// TIA Portal V15.1 program export: 1 tag tables, 0 data types, 3 data blocks, 7 code blocks (in call order from the OBs), 3 instance data blocks

VAR_GLOBAL   // PLC tag table "IO"
   PSH_101 AT %I0.0 : Bool;   // Scrubber high pressure
   LSH_102 AT %I0.1 : Bool;   // Scrubber high level
   LSHH_103 AT %I0.2 : Bool;   // Scrubber high-high level
   BR01_Run AT %I0.3 : Bool;   // BR01 run feedback
   S1_BR01_Start AT %I0.4 : Bool;   // BR01 START push button
   BR01_Fault AT %I0.5 : Bool;   // BR01 fault (lockout)
   S3_BR01_Stop AT %I0.6 : Bool;   // BR01 STOP push button
   S0_EStopStatus AT %I1.0 : Bool;   // E-STOP status (NC1)
   S2_FaultReset AT %I1.1 : Bool;   // FAULT RESET push button
   LSL_TK01 AT %I1.2 : Bool;   // TK01 low level
   LSL_TK02 AT %I1.3 : Bool;   // TK02 low level
   BR02_Run AT %I1.4 : Bool;   // BR02 run feedback
   BR02_Fault AT %I1.5 : Bool;   // BR02 fault (lockout)
   Rfuel2_BR02_DieselMode AT %I12.0 : Bool;   // BR02 diesel mode
   S4_BR01_Auto AT %I12.1 : Bool;   // BR01 AUTO/MAN selector (closed = AUTO)
   S5_BR02_Auto AT %I12.2 : Bool;   // BR02 AUTO/MAN selector (closed = AUTO)
   S6_BR02_Start AT %I12.3 : Bool;   // BR02 START push button
   S7_BR02_Stop AT %I12.4 : Bool;   // BR02 STOP push button
   BR01_TL_Cmd AT %Q0.0 : Bool;   // BR01 heat request (TL) + H1 1st stage lamp
   BR01_TR_Cmd AT %Q0.1 : Bool;   // BR01 2nd stage (TR) + H2 2nd stage lamp
   XV_401_Cmd AT %Q0.2 : Bool;   // XV-401 Flare SV (NO)
   XV_402_Cmd AT %Q0.3 : Bool;   // XV-402 Drain SV (NC)
   XV_403_Cmd AT %Q0.4 : Bool;   // XV-403 Suction SV (NC)
   BR02_L_Cmd AT %Q0.5 : Bool;   // BR02 start (L)
   BR02_T2_Cmd AT %Q0.6 : Bool;   // BR02 high fire (T2)
   BR02_Stage1Lamp_Cmd AT %Q0.7 : Bool;   // BR02 1st stage lamp H5
   BR02_Stage2Lamp_Cmd AT %Q1.0 : Bool;   // BR02 2nd stage lamp H6
   TE_501_Raw AT %IW96 : Int;   // TK01 inlet oil temperature
   TE_502_Raw AT %IW98 : Int;   // TK01 outlet oil temperature
   TE_503_Raw AT %IW100 : Int;   // TK02 inlet oil temperature
   TE_504_Raw AT %IW102 : Int;   // TK02 outlet oil temperature
END_VAR

DATA_BLOCK "HmiAlm"   // DB6
{ S7_Optimized_Access := 'TRUE' }
VERSION : 0.1
// stored: AutoNumber false, MemoryReserve 100
   VAR
      Common : Word;   // 0007 / H-05: x0 E-STOP active or not reset [C01]; x1 Scrubber trip: high pressure PSH-101 [C03 / C06a (PH proposal: cause memory)]; x2 Scrubber trip: high-high level LSHH-103 [C05 / C06a (PH proposal: cause memory)]; x3 Scrubber held after power-up: RESET required [S-01 / C06a (PH proposal)]; x4 Scrubber high level LSH-102 [C04 (Client)]; x5 Setting rejected: out of range [R-11]; x6 Scrubber drain open too long: drain closed [C04a]; x7 LSH-102 fault: LSHH-103 without LSH-102 [C04b]
      BR01 : Word;   // 0007 / H-05: x0 BR01 stopped by E-STOP: RESET + START [C01]; x1 BR01 thermocouple fault [C07d]; x2 BR01 burner lockout [C07e]; x3 BR01 failed to start [C07f]; x4 BR01 stopped by itself [C07g]; x5 BR01 RUN without request [R-09]; x6 TK01 level low: burner held [C07a (PH proposal: alarm; Client: permissive)]
      BR02 : Word;   // 0007 / H-05: x0 BR02 stopped by E-STOP: RESET + START [C01]; x1 BR02 thermocouple fault [C08d]; x2 BR02 burner lockout [C08e]; x3 BR02 failed to start [C08f]; x4 BR02 stopped by itself [C08g]; x5 BR02 RUN without request [R-09]; x6 TK02 level low: burner held [C08a (PH proposal: alarm; Client: permissive)]
   END_VAR
BEGIN
END_DATA_BLOCK

DATA_BLOCK "Par"   // DB1
{ S7_Optimized_Access := 'TRUE' }
VERSION : 0.1
// stored: AutoNumber false, MemoryReserve 100
   VAR RETAIN
      SP : Int := 700;   // HMI entry: Setpoint, 0.1 degC (C07b)
      HYST : Int := 50;   // HMI entry: Restart hysteresis, 0.1 degC (C07b)
      STG : Int := 100;   // HMI entry: 2nd stage below SP - STG, 0.1 degC (C07c)
      TStart : Time := T#2M;   // HMI entry: Max. time heat request -> RUN (C07f)
      TDrnOn : Time := T#3S;   // HMI entry: Scrubber high level before drain opens (C04)
      TDrnOff : Time := T#5S;   // HMI entry: Scrubber level gone before drain closes (C04)
      TDrnMax : Time := T#10M;   // HMI entry: Scrubber drain max. continuous open time (C04a)
      SP_V : Int := 700;   // Validated value used by the program (R-11)
      HYST_V : Int := 50;   // Validated value used by the program (R-11)
      STG_V : Int := 100;   // Validated value used by the program (R-11)
      TStart_V : Time := T#2M;   // Validated value used by the program (R-11)
      TDrnOn_V : Time := T#3S;   // Validated value used by the program (R-11)
      TDrnOff_V : Time := T#5S;   // Validated value used by the program (R-11)
      TDrnMax_V : Time := T#10M;   // Validated value used by the program (R-11)
   END_VAR
BEGIN
END_DATA_BLOCK

DATA_BLOCK "Sys"   // DB2
{ S7_Optimized_Access := 'TRUE' }
VERSION : 0.1
// stored: AutoNumber false, MemoryReserve 100
   VAR
      FirstScan : Bool;   // Set by OB100, cleared at the end of Main (C02)
      EStopOK : Bool;   // E-STOP latch: 1 = released and RESET given (C01)
      ResetPulse : Bool;   // RESET S2 rising edge, one scan (R-06)
      ResetMem : Bool;   // RESET edge memory (R-06)
      Alm_EStop : Bool;   // HMI alarm: E-STOP (C01)
      Alm_ParRejected : Bool;   // HMI alarm: a parameter entry was out of range (R-11)
   END_VAR
BEGIN
END_DATA_BLOCK

ORGANIZATION_BLOCK "Main"   // OB1, LAD, ProgramCycle
TITLE = Main
{ S7_Optimized_Access := 'TRUE' }
VERSION : 0.1
// Calls the blocks in a fixed order; no logic here (decisions/0006)
// stored: AutoNumber false, IsIECCheckEnabled false, SetENOAutomatically False
   VAR_INPUT
      Initial_Call : Bool;
      Remanence : Bool;
   END_VAR
BEGIN

REGION Network 1: decisions/0006 — Common: E-STOP latch, RESET edge, parameters
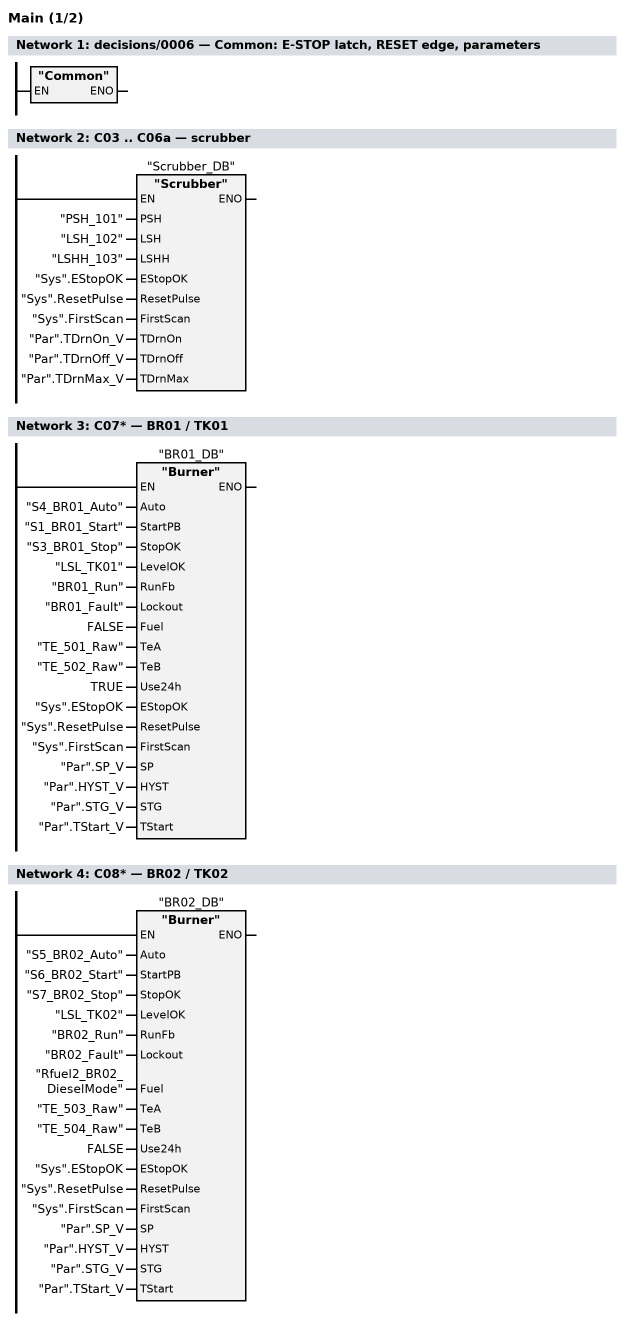
   RUNG wire#powerrail
      "Common"()
   END_RUNG
   // the same network as SCL:
   "Common"();
END_REGION

REGION Network 2: C03 .. C06a — scrubber
   RUNG wire#powerrail
      "Scrubber_DB"(PSH := "PSH_101", LSH := "LSH_102", LSHH := "LSHH_103", EStopOK := "Sys".EStopOK, ResetPulse := "Sys".ResetPulse, FirstScan := "Sys".FirstScan, TDrnOn := "Par".TDrnOn_V, TDrnOff := "Par".TDrnOff_V, TDrnMax := "Par".TDrnMax_V)
   END_RUNG
   // the same network as SCL:
   "Scrubber_DB"(PSH := "PSH_101",   // "Scrubber"
                 LSH := "LSH_102",
                 LSHH := "LSHH_103",
                 EStopOK := "Sys".EStopOK,
                 ResetPulse := "Sys".ResetPulse,
                 FirstScan := "Sys".FirstScan,
                 TDrnOn := "Par".TDrnOn_V,
                 TDrnOff := "Par".TDrnOff_V,
                 TDrnMax := "Par".TDrnMax_V);
END_REGION

REGION Network 3: C07* — BR01 / TK01
   RUNG wire#powerrail
      "BR01_DB"(Auto := "S4_BR01_Auto", StartPB := "S1_BR01_Start", StopOK := "S3_BR01_Stop", LevelOK := "LSL_TK01", RunFb := "BR01_Run", Lockout := "BR01_Fault", Fuel := FALSE, TeA := "TE_501_Raw", TeB := "TE_502_Raw", Use24h := TRUE, EStopOK := "Sys".EStopOK, ResetPulse := "Sys".ResetPulse, FirstScan := "Sys".FirstScan, SP := "Par".SP_V, HYST := "Par".HYST_V, STG := "Par".STG_V, TStart := "Par".TStart_V)
   END_RUNG
   // the same network as SCL:
   "BR01_DB"(Auto := "S4_BR01_Auto",   // "Burner"
             StartPB := "S1_BR01_Start",
             StopOK := "S3_BR01_Stop",
             LevelOK := "LSL_TK01",
             RunFb := "BR01_Run",
             Lockout := "BR01_Fault",
             Fuel := FALSE,
             TeA := "TE_501_Raw",
             TeB := "TE_502_Raw",
             Use24h := TRUE,
             EStopOK := "Sys".EStopOK,
             ResetPulse := "Sys".ResetPulse,
             FirstScan := "Sys".FirstScan,
             SP := "Par".SP_V,
             HYST := "Par".HYST_V,
             STG := "Par".STG_V,
             TStart := "Par".TStart_V);
END_REGION

REGION Network 4: C08* — BR02 / TK02
   RUNG wire#powerrail
      "BR02_DB"(Auto := "S5_BR02_Auto", StartPB := "S6_BR02_Start", StopOK := "S7_BR02_Stop", LevelOK := "LSL_TK02", RunFb := "BR02_Run", Lockout := "BR02_Fault", Fuel := "Rfuel2_BR02_DieselMode", TeA := "TE_503_Raw", TeB := "TE_504_Raw", Use24h := FALSE, EStopOK := "Sys".EStopOK, ResetPulse := "Sys".ResetPulse, FirstScan := "Sys".FirstScan, SP := "Par".SP_V, HYST := "Par".HYST_V, STG := "Par".STG_V, TStart := "Par".TStart_V)
   END_RUNG
   // the same network as SCL:
   "BR02_DB"(Auto := "S5_BR02_Auto",   // "Burner"
             StartPB := "S6_BR02_Start",
             StopOK := "S7_BR02_Stop",
             LevelOK := "LSL_TK02",
             RunFb := "BR02_Run",
             Lockout := "BR02_Fault",
             Fuel := "Rfuel2_BR02_DieselMode",
             TeA := "TE_503_Raw",
             TeB := "TE_504_Raw",
             Use24h := FALSE,
             EStopOK := "Sys".EStopOK,
             ResetPulse := "Sys".ResetPulse,
             FirstScan := "Sys".FirstScan,
             SP := "Par".SP_V,
             HYST := "Par".HYST_V,
             STG := "Par".STG_V,
             TStart := "Par".TStart_V);
END_REGION

REGION Network 5: E1 .. E7 — outputs
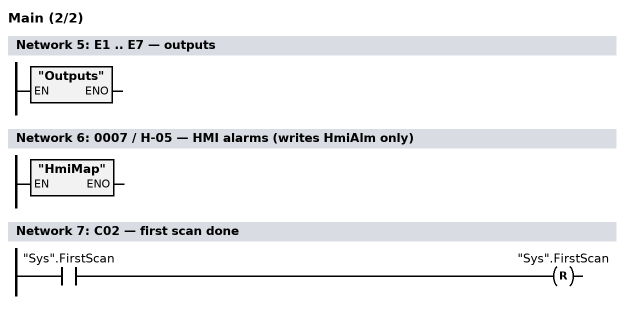
   RUNG wire#powerrail
      "Outputs"()
   END_RUNG
   // the same network as SCL:
   "Outputs"();
END_REGION

REGION Network 6: 0007 / H-05 — HMI alarms (writes HmiAlm only)
   RUNG wire#powerrail
      "HmiMap"()
   END_RUNG
   // the same network as SCL:
   "HmiMap"();
END_REGION

REGION Network 7: C02 — first scan done
   RUNG wire#powerrail
      Contact( "Sys".FirstScan )
      R_Coil( "Sys".FirstScan )
   END_RUNG
   // the same network as SCL:
   IF "Sys".FirstScan THEN "Sys".FirstScan := FALSE; END_IF;
END_REGION
END_ORGANIZATION_BLOCK

FUNCTION "Common" : Void   // FC1, LAD
TITLE = Common
{ S7_Optimized_Access := 'TRUE' }
VERSION : 0.1
// E-STOP latch, RESET edge, parameter check (decisions/0006)
// stored: AutoNumber false, IsIECCheckEnabled false, SetENOAutomatically False
   VAR_TEMP   // added for the SCL form of the ladder/FBD networks
      _w1 : Bool;
   END_VAR
BEGIN

REGION Network 1: R-06 — RESET edge (not on first scan)
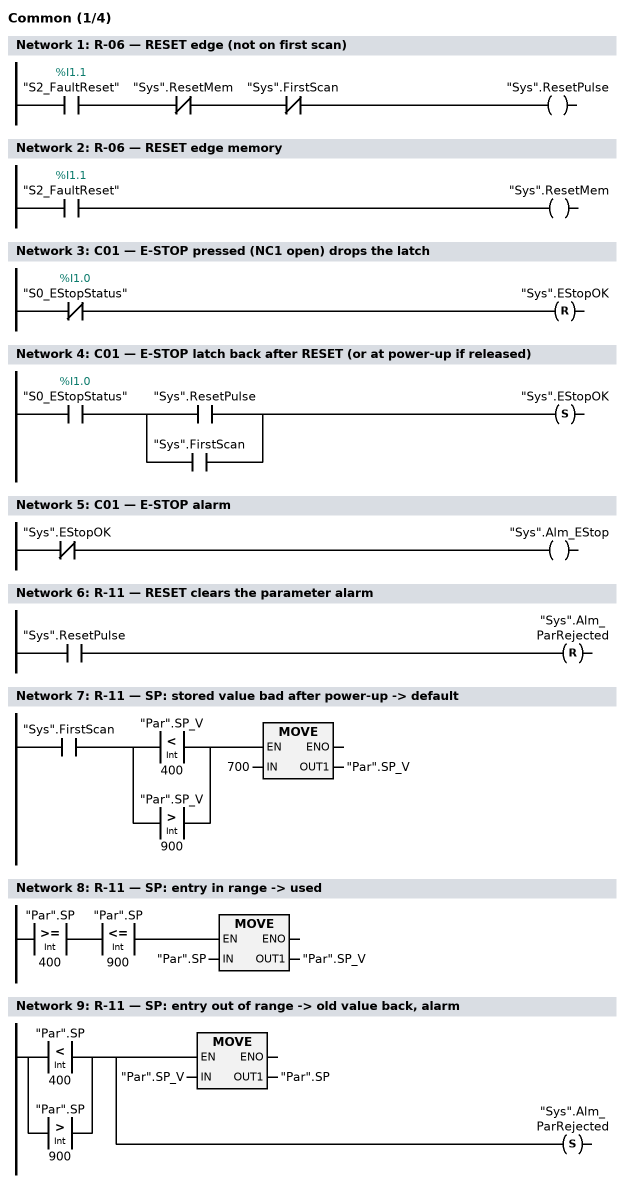
   RUNG wire#powerrail
      Contact( "S2_FaultReset" )
      I_Contact( "Sys".ResetMem )
      I_Contact( "Sys".FirstScan )
      Coil( "Sys".ResetPulse )
   END_RUNG
   // the same network as SCL:
   "Sys".ResetPulse := "S2_FaultReset" AND NOT "Sys".ResetMem AND NOT "Sys".FirstScan;
END_REGION

REGION Network 2: R-06 — RESET edge memory
   RUNG wire#powerrail
      Contact( "S2_FaultReset" )
      Coil( "Sys".ResetMem )
   END_RUNG
   // the same network as SCL:
   "Sys".ResetMem := "S2_FaultReset";
END_REGION

REGION Network 3: C01 — E-STOP pressed (NC1 open) drops the latch
   RUNG wire#powerrail
      I_Contact( "S0_EStopStatus" )
      R_Coil( "Sys".EStopOK )
   END_RUNG
   // the same network as SCL:
   IF NOT "S0_EStopStatus" THEN "Sys".EStopOK := FALSE; END_IF;
END_REGION

REGION Network 4: C01 — E-STOP latch back after RESET (or at power-up if released)
   RUNG wire#powerrail
      Contact( "S0_EStopStatus" )
      wire#w1
      Contact( "Sys".ResetPulse )
      wire#w2
      S_Coil( "Sys".EStopOK )
   END_RUNG
   RUNG wire#w1
      Contact( "Sys".FirstScan )
   END_RUNG wire#w2
   // the same network as SCL:
   IF "S0_EStopStatus" AND ("Sys".ResetPulse OR "Sys".FirstScan) THEN "Sys".EStopOK := TRUE; END_IF;
END_REGION

REGION Network 5: C01 — E-STOP alarm
   RUNG wire#powerrail
      I_Contact( "Sys".EStopOK )
      Coil( "Sys".Alm_EStop )
   END_RUNG
   // the same network as SCL:
   "Sys".Alm_EStop := NOT "Sys".EStopOK;
END_REGION

REGION Network 6: R-11 — RESET clears the parameter alarm
   RUNG wire#powerrail
      Contact( "Sys".ResetPulse )
      R_Coil( "Sys".Alm_ParRejected )
   END_RUNG
   // the same network as SCL:
   IF "Sys".ResetPulse THEN "Sys".Alm_ParRejected := FALSE; END_IF;
END_REGION

REGION Network 7: R-11 — SP: stored value bad after power-up -> default
   RUNG wire#powerrail
      Contact( "Sys".FirstScan )
      wire#w1
      { S7_Templates := "SrcType := Int" } LT_Contact(in1 := "Par".SP_V, in2 := 400)
      wire#w2
      { S7_GenerateENO := "TRUE" } Move(in := 700, out1 => "Par".SP_V)
   END_RUNG
   RUNG wire#w1
      { S7_Templates := "SrcType := Int" } GT_Contact(in1 := "Par".SP_V, in2 := 900)
   END_RUNG wire#w2
   // the same network as SCL:
   IF "Sys".FirstScan AND (("Par".SP_V < 400) OR ("Par".SP_V > 900)) THEN "Par".SP_V := 700; END_IF;
END_REGION

REGION Network 8: R-11 — SP: entry in range -> used
   RUNG wire#powerrail
      { S7_Templates := "SrcType := Int" } GE_Contact(in1 := "Par".SP, in2 := 400)
      { S7_Templates := "SrcType := Int" } LE_Contact(in1 := "Par".SP, in2 := 900)
      { S7_GenerateENO := "TRUE" } Move(in := "Par".SP, out1 => "Par".SP_V)
   END_RUNG
   // the same network as SCL:
   IF ("Par".SP >= 400) AND ("Par".SP <= 900) THEN "Par".SP_V := "Par".SP; END_IF;
END_REGION

REGION Network 9: R-11 — SP: entry out of range -> old value back, alarm
   RUNG wire#powerrail
      { S7_Templates := "SrcType := Int" } LT_Contact(in1 := "Par".SP, in2 := 400)
      wire#w1
      { S7_GenerateENO := "TRUE" } Move(in := "Par".SP_V, out1 => "Par".SP)
   END_RUNG
   RUNG wire#powerrail
      { S7_Templates := "SrcType := Int" } GT_Contact(in1 := "Par".SP, in2 := 900)
   END_RUNG wire#w1
   RUNG wire#w1
      S_Coil( "Sys".Alm_ParRejected )
   END_RUNG
   // the same network as SCL:
   #_w1 := ("Par".SP < 400) OR ("Par".SP > 900);
   IF #_w1 THEN
       "Par".SP := "Par".SP_V;
       "Sys".Alm_ParRejected := TRUE;
   END_IF;
END_REGION

REGION Network 10: R-11 — HYST: stored value bad after power-up -> default
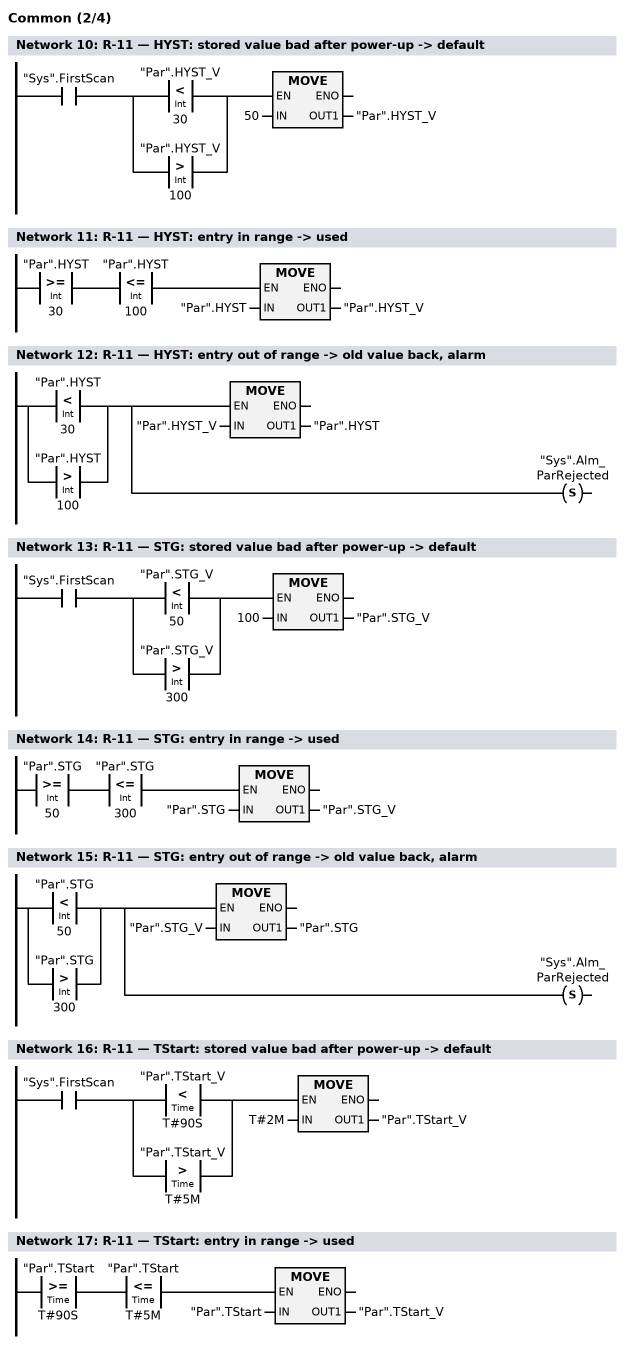
   RUNG wire#powerrail
      Contact( "Sys".FirstScan )
      wire#w1
      { S7_Templates := "SrcType := Int" } LT_Contact(in1 := "Par".HYST_V, in2 := 30)
      wire#w2
      { S7_GenerateENO := "TRUE" } Move(in := 50, out1 => "Par".HYST_V)
   END_RUNG
   RUNG wire#w1
      { S7_Templates := "SrcType := Int" } GT_Contact(in1 := "Par".HYST_V, in2 := 100)
   END_RUNG wire#w2
   // the same network as SCL:
   IF "Sys".FirstScan AND (("Par".HYST_V < 30) OR ("Par".HYST_V > 100)) THEN "Par".HYST_V := 50; END_IF;
END_REGION

REGION Network 11: R-11 — HYST: entry in range -> used
   RUNG wire#powerrail
      { S7_Templates := "SrcType := Int" } GE_Contact(in1 := "Par".HYST, in2 := 30)
      { S7_Templates := "SrcType := Int" } LE_Contact(in1 := "Par".HYST, in2 := 100)
      { S7_GenerateENO := "TRUE" } Move(in := "Par".HYST, out1 => "Par".HYST_V)
   END_RUNG
   // the same network as SCL:
   IF ("Par".HYST >= 30) AND ("Par".HYST <= 100) THEN "Par".HYST_V := "Par".HYST; END_IF;
END_REGION

REGION Network 12: R-11 — HYST: entry out of range -> old value back, alarm
   RUNG wire#powerrail
      { S7_Templates := "SrcType := Int" } LT_Contact(in1 := "Par".HYST, in2 := 30)
      wire#w1
      { S7_GenerateENO := "TRUE" } Move(in := "Par".HYST_V, out1 => "Par".HYST)
   END_RUNG
   RUNG wire#powerrail
      { S7_Templates := "SrcType := Int" } GT_Contact(in1 := "Par".HYST, in2 := 100)
   END_RUNG wire#w1
   RUNG wire#w1
      S_Coil( "Sys".Alm_ParRejected )
   END_RUNG
   // the same network as SCL:
   #_w1 := ("Par".HYST < 30) OR ("Par".HYST > 100);
   IF #_w1 THEN
       "Par".HYST := "Par".HYST_V;
       "Sys".Alm_ParRejected := TRUE;
   END_IF;
END_REGION

REGION Network 13: R-11 — STG: stored value bad after power-up -> default
   RUNG wire#powerrail
      Contact( "Sys".FirstScan )
      wire#w1
      { S7_Templates := "SrcType := Int" } LT_Contact(in1 := "Par".STG_V, in2 := 50)
      wire#w2
      { S7_GenerateENO := "TRUE" } Move(in := 100, out1 => "Par".STG_V)
   END_RUNG
   RUNG wire#w1
      { S7_Templates := "SrcType := Int" } GT_Contact(in1 := "Par".STG_V, in2 := 300)
   END_RUNG wire#w2
   // the same network as SCL:
   IF "Sys".FirstScan AND (("Par".STG_V < 50) OR ("Par".STG_V > 300)) THEN "Par".STG_V := 100; END_IF;
END_REGION

REGION Network 14: R-11 — STG: entry in range -> used
   RUNG wire#powerrail
      { S7_Templates := "SrcType := Int" } GE_Contact(in1 := "Par".STG, in2 := 50)
      { S7_Templates := "SrcType := Int" } LE_Contact(in1 := "Par".STG, in2 := 300)
      { S7_GenerateENO := "TRUE" } Move(in := "Par".STG, out1 => "Par".STG_V)
   END_RUNG
   // the same network as SCL:
   IF ("Par".STG >= 50) AND ("Par".STG <= 300) THEN "Par".STG_V := "Par".STG; END_IF;
END_REGION

REGION Network 15: R-11 — STG: entry out of range -> old value back, alarm
   RUNG wire#powerrail
      { S7_Templates := "SrcType := Int" } LT_Contact(in1 := "Par".STG, in2 := 50)
      wire#w1
      { S7_GenerateENO := "TRUE" } Move(in := "Par".STG_V, out1 => "Par".STG)
   END_RUNG
   RUNG wire#powerrail
      { S7_Templates := "SrcType := Int" } GT_Contact(in1 := "Par".STG, in2 := 300)
   END_RUNG wire#w1
   RUNG wire#w1
      S_Coil( "Sys".Alm_ParRejected )
   END_RUNG
   // the same network as SCL:
   #_w1 := ("Par".STG < 50) OR ("Par".STG > 300);
   IF #_w1 THEN
       "Par".STG := "Par".STG_V;
       "Sys".Alm_ParRejected := TRUE;
   END_IF;
END_REGION

REGION Network 16: R-11 — TStart: stored value bad after power-up -> default
   RUNG wire#powerrail
      Contact( "Sys".FirstScan )
      wire#w1
      { S7_Templates := "SrcType := Time" } LT_Contact(in1 := "Par".TStart_V, in2 := T#90S)
      wire#w2
      { S7_GenerateENO := "TRUE" } Move(in := T#2M, out1 => "Par".TStart_V)
   END_RUNG
   RUNG wire#w1
      { S7_Templates := "SrcType := Time" } GT_Contact(in1 := "Par".TStart_V, in2 := T#5M)
   END_RUNG wire#w2
   // the same network as SCL:
   IF "Sys".FirstScan AND (("Par".TStart_V < T#90S) OR ("Par".TStart_V > T#5M)) THEN
       "Par".TStart_V := T#2M;
   END_IF;
END_REGION

REGION Network 17: R-11 — TStart: entry in range -> used
   RUNG wire#powerrail
      { S7_Templates := "SrcType := Time" } GE_Contact(in1 := "Par".TStart, in2 := T#90S)
      { S7_Templates := "SrcType := Time" } LE_Contact(in1 := "Par".TStart, in2 := T#5M)
      { S7_GenerateENO := "TRUE" } Move(in := "Par".TStart, out1 => "Par".TStart_V)
   END_RUNG
   // the same network as SCL:
   IF ("Par".TStart >= T#90S) AND ("Par".TStart <= T#5M) THEN "Par".TStart_V := "Par".TStart; END_IF;
END_REGION

REGION Network 18: R-11 — TStart: entry out of range -> old value back, alarm
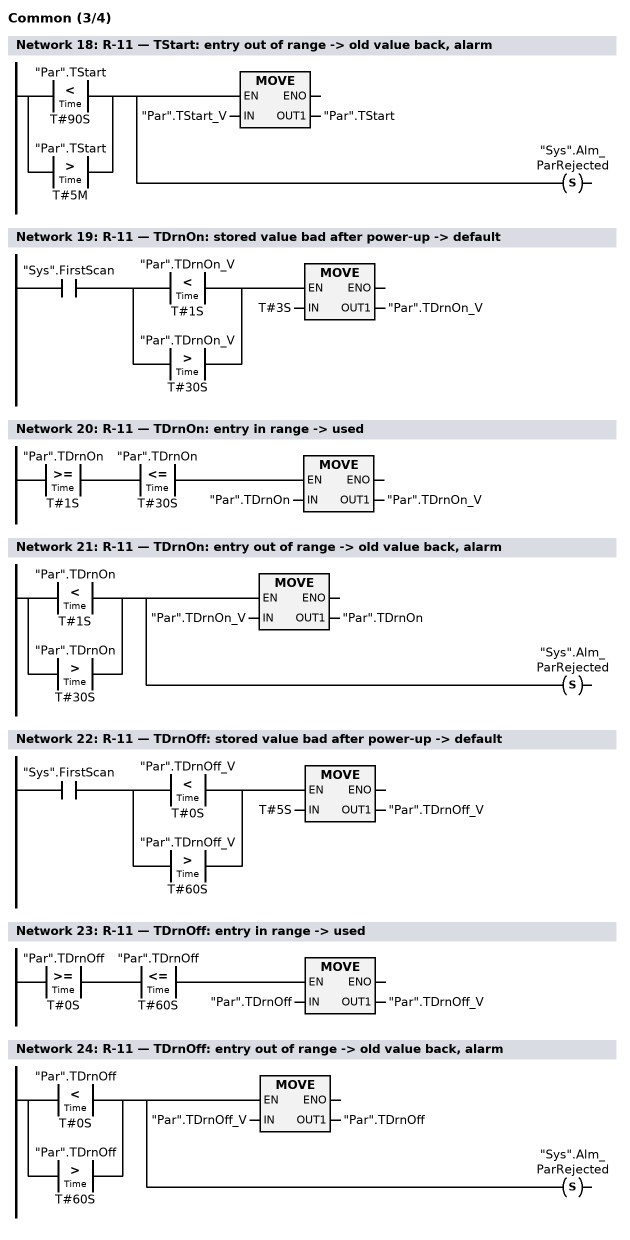
   RUNG wire#powerrail
      { S7_Templates := "SrcType := Time" } LT_Contact(in1 := "Par".TStart, in2 := T#90S)
      wire#w1
      { S7_GenerateENO := "TRUE" } Move(in := "Par".TStart_V, out1 => "Par".TStart)
   END_RUNG
   RUNG wire#powerrail
      { S7_Templates := "SrcType := Time" } GT_Contact(in1 := "Par".TStart, in2 := T#5M)
   END_RUNG wire#w1
   RUNG wire#w1
      S_Coil( "Sys".Alm_ParRejected )
   END_RUNG
   // the same network as SCL:
   #_w1 := ("Par".TStart < T#90S) OR ("Par".TStart > T#5M);
   IF #_w1 THEN
       "Par".TStart := "Par".TStart_V;
       "Sys".Alm_ParRejected := TRUE;
   END_IF;
END_REGION

REGION Network 19: R-11 — TDrnOn: stored value bad after power-up -> default
   RUNG wire#powerrail
      Contact( "Sys".FirstScan )
      wire#w1
      { S7_Templates := "SrcType := Time" } LT_Contact(in1 := "Par".TDrnOn_V, in2 := T#1S)
      wire#w2
      { S7_GenerateENO := "TRUE" } Move(in := T#3S, out1 => "Par".TDrnOn_V)
   END_RUNG
   RUNG wire#w1
      { S7_Templates := "SrcType := Time" } GT_Contact(in1 := "Par".TDrnOn_V, in2 := T#30S)
   END_RUNG wire#w2
   // the same network as SCL:
   IF "Sys".FirstScan AND (("Par".TDrnOn_V < T#1S) OR ("Par".TDrnOn_V > T#30S)) THEN
       "Par".TDrnOn_V := T#3S;
   END_IF;
END_REGION

REGION Network 20: R-11 — TDrnOn: entry in range -> used
   RUNG wire#powerrail
      { S7_Templates := "SrcType := Time" } GE_Contact(in1 := "Par".TDrnOn, in2 := T#1S)
      { S7_Templates := "SrcType := Time" } LE_Contact(in1 := "Par".TDrnOn, in2 := T#30S)
      { S7_GenerateENO := "TRUE" } Move(in := "Par".TDrnOn, out1 => "Par".TDrnOn_V)
   END_RUNG
   // the same network as SCL:
   IF ("Par".TDrnOn >= T#1S) AND ("Par".TDrnOn <= T#30S) THEN "Par".TDrnOn_V := "Par".TDrnOn; END_IF;
END_REGION

REGION Network 21: R-11 — TDrnOn: entry out of range -> old value back, alarm
   RUNG wire#powerrail
      { S7_Templates := "SrcType := Time" } LT_Contact(in1 := "Par".TDrnOn, in2 := T#1S)
      wire#w1
      { S7_GenerateENO := "TRUE" } Move(in := "Par".TDrnOn_V, out1 => "Par".TDrnOn)
   END_RUNG
   RUNG wire#powerrail
      { S7_Templates := "SrcType := Time" } GT_Contact(in1 := "Par".TDrnOn, in2 := T#30S)
   END_RUNG wire#w1
   RUNG wire#w1
      S_Coil( "Sys".Alm_ParRejected )
   END_RUNG
   // the same network as SCL:
   #_w1 := ("Par".TDrnOn < T#1S) OR ("Par".TDrnOn > T#30S);
   IF #_w1 THEN
       "Par".TDrnOn := "Par".TDrnOn_V;
       "Sys".Alm_ParRejected := TRUE;
   END_IF;
END_REGION

REGION Network 22: R-11 — TDrnOff: stored value bad after power-up -> default
   RUNG wire#powerrail
      Contact( "Sys".FirstScan )
      wire#w1
      { S7_Templates := "SrcType := Time" } LT_Contact(in1 := "Par".TDrnOff_V, in2 := T#0S)
      wire#w2
      { S7_GenerateENO := "TRUE" } Move(in := T#5S, out1 => "Par".TDrnOff_V)
   END_RUNG
   RUNG wire#w1
      { S7_Templates := "SrcType := Time" } GT_Contact(in1 := "Par".TDrnOff_V, in2 := T#60S)
   END_RUNG wire#w2
   // the same network as SCL:
   IF "Sys".FirstScan AND (("Par".TDrnOff_V < T#0S) OR ("Par".TDrnOff_V > T#60S)) THEN
       "Par".TDrnOff_V := T#5S;
   END_IF;
END_REGION

REGION Network 23: R-11 — TDrnOff: entry in range -> used
   RUNG wire#powerrail
      { S7_Templates := "SrcType := Time" } GE_Contact(in1 := "Par".TDrnOff, in2 := T#0S)
      { S7_Templates := "SrcType := Time" } LE_Contact(in1 := "Par".TDrnOff, in2 := T#60S)
      { S7_GenerateENO := "TRUE" } Move(in := "Par".TDrnOff, out1 => "Par".TDrnOff_V)
   END_RUNG
   // the same network as SCL:
   IF ("Par".TDrnOff >= T#0S) AND ("Par".TDrnOff <= T#60S) THEN "Par".TDrnOff_V := "Par".TDrnOff; END_IF;
END_REGION

REGION Network 24: R-11 — TDrnOff: entry out of range -> old value back, alarm
   RUNG wire#powerrail
      { S7_Templates := "SrcType := Time" } LT_Contact(in1 := "Par".TDrnOff, in2 := T#0S)
      wire#w1
      { S7_GenerateENO := "TRUE" } Move(in := "Par".TDrnOff_V, out1 => "Par".TDrnOff)
   END_RUNG
   RUNG wire#powerrail
      { S7_Templates := "SrcType := Time" } GT_Contact(in1 := "Par".TDrnOff, in2 := T#60S)
   END_RUNG wire#w1
   RUNG wire#w1
      S_Coil( "Sys".Alm_ParRejected )
   END_RUNG
   // the same network as SCL:
   #_w1 := ("Par".TDrnOff < T#0S) OR ("Par".TDrnOff > T#60S);
   IF #_w1 THEN
       "Par".TDrnOff := "Par".TDrnOff_V;
       "Sys".Alm_ParRejected := TRUE;
   END_IF;
END_REGION

REGION Network 25: R-11 — TDrnMax: stored value bad after power-up -> default
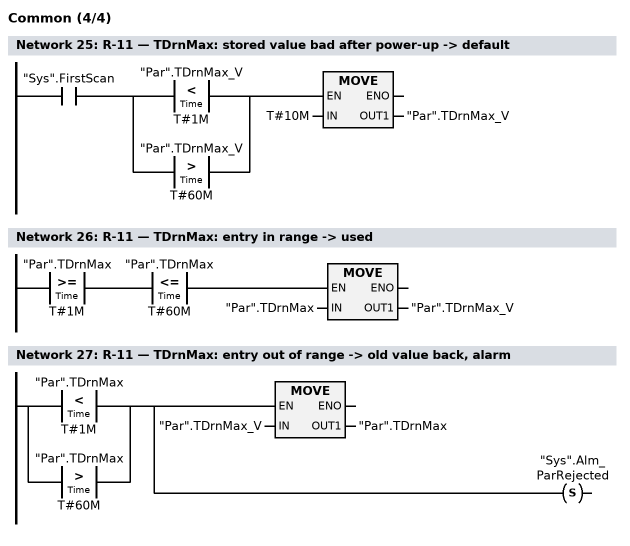
   RUNG wire#powerrail
      Contact( "Sys".FirstScan )
      wire#w1
      { S7_Templates := "SrcType := Time" } LT_Contact(in1 := "Par".TDrnMax_V, in2 := T#1M)
      wire#w2
      { S7_GenerateENO := "TRUE" } Move(in := T#10M, out1 => "Par".TDrnMax_V)
   END_RUNG
   RUNG wire#w1
      { S7_Templates := "SrcType := Time" } GT_Contact(in1 := "Par".TDrnMax_V, in2 := T#60M)
   END_RUNG wire#w2
   // the same network as SCL:
   IF "Sys".FirstScan AND (("Par".TDrnMax_V < T#1M) OR ("Par".TDrnMax_V > T#60M)) THEN
       "Par".TDrnMax_V := T#10M;
   END_IF;
END_REGION

REGION Network 26: R-11 — TDrnMax: entry in range -> used
   RUNG wire#powerrail
      { S7_Templates := "SrcType := Time" } GE_Contact(in1 := "Par".TDrnMax, in2 := T#1M)
      { S7_Templates := "SrcType := Time" } LE_Contact(in1 := "Par".TDrnMax, in2 := T#60M)
      { S7_GenerateENO := "TRUE" } Move(in := "Par".TDrnMax, out1 => "Par".TDrnMax_V)
   END_RUNG
   // the same network as SCL:
   IF ("Par".TDrnMax >= T#1M) AND ("Par".TDrnMax <= T#60M) THEN "Par".TDrnMax_V := "Par".TDrnMax; END_IF;
END_REGION

REGION Network 27: R-11 — TDrnMax: entry out of range -> old value back, alarm
   RUNG wire#powerrail
      { S7_Templates := "SrcType := Time" } LT_Contact(in1 := "Par".TDrnMax, in2 := T#1M)
      wire#w1
      { S7_GenerateENO := "TRUE" } Move(in := "Par".TDrnMax_V, out1 => "Par".TDrnMax)
   END_RUNG
   RUNG wire#powerrail
      { S7_Templates := "SrcType := Time" } GT_Contact(in1 := "Par".TDrnMax, in2 := T#60M)
   END_RUNG wire#w1
   RUNG wire#w1
      S_Coil( "Sys".Alm_ParRejected )
   END_RUNG
   // the same network as SCL:
   #_w1 := ("Par".TDrnMax < T#1M) OR ("Par".TDrnMax > T#60M);
   IF #_w1 THEN
       "Par".TDrnMax := "Par".TDrnMax_V;
       "Sys".Alm_ParRejected := TRUE;
   END_IF;
END_REGION
END_FUNCTION

FUNCTION_BLOCK "Scrubber"   // FB2, LAD
TITLE = Scrubber
{ S7_Optimized_Access := 'TRUE' }
VERSION : 0.1
// Gas scrubber, docs/التشغيل.md §1
// stored: AutoNumber false, IsIECCheckEnabled false, MemoryReserve 100, SetENOAutomatically False
   VAR_INPUT
      PSH : Bool;   // PSH-101 healthy (contact closed)
      LSH : Bool;   // LSH-102 healthy
      LSHH : Bool;   // LSHH-103 healthy
      EStopOK : Bool;   // Sys.EStopOK
      ResetPulse : Bool;   // Sys.ResetPulse
      FirstScan : Bool;   // Sys.FirstScan
      TDrnOn : Time;   // Par.TDrnOn_V (C04)
      TDrnOff : Time;   // Par.TDrnOff_V (C04)
      TDrnMax : Time;   // Par.TDrnMax_V (C04a)
   END_VAR
   VAR_OUTPUT
      Tripped : Bool;   // Suction trip latch C01/C02/C03/C05: XV-403 closed until RESET
      FlareTrip : Bool;   // Flare trip latch C01/C02/C03: XV-401 open until RESET
      ValvesNormal : Bool;   // No trip latched: flare closed and suction open (HMI)
      FlareCmd : Bool;   // Q0.2 XV-401 (NO): 1 = energised = closed
      DrainCmd : Bool;   // Q0.3 XV-402 (NC): 1 = energised = open (C04 / C05)
      SuctionCmd : Bool;   // Q0.4 XV-403 (NC): 1 = energised = open
      F_DrainTO : Bool;   // C04a: drain open too long, latched until RESET
      F_LshFault : Bool;   // C04b: LSHH-103 without LSH-102, latched until RESET
      Alm_PSH : Bool;   // HMI alarm C03
      Alm_LSH : Bool;   // HMI alarm C04
      Alm_LSHH : Bool;   // HMI alarm C05
      Cause_EStop : Bool;   // C06a / F44: E-STOP cause, latched until healthy RESET
      Cause_PSH : Bool;   // C06a / F44: PSH-101 cause, latched until healthy RESET
      Cause_LSHH : Bool;   // C06a / F44: LSHH-103 cause, latched until healthy RESET
      Cause_PwrUp : Bool;   // C06a / F44: power-up cause, latched until healthy RESET
      FirstOut : Int;   // C06a / 0007 D5: 0 none, 1 E-STOP, 2 PSH, 3 LSHH, 4 power-up
   END_VAR
   VAR
      LevelHigh : Bool;
      DrnDemand : Bool;
      T_DrnOn : TON_TIME;
      T_DrnOff : TON_TIME;
      T_DrnMax : TON_TIME;
      T_LshFlt : TON_TIME;
   END_VAR
BEGIN

REGION Network 1: C04 — LSH-102 high level alarm
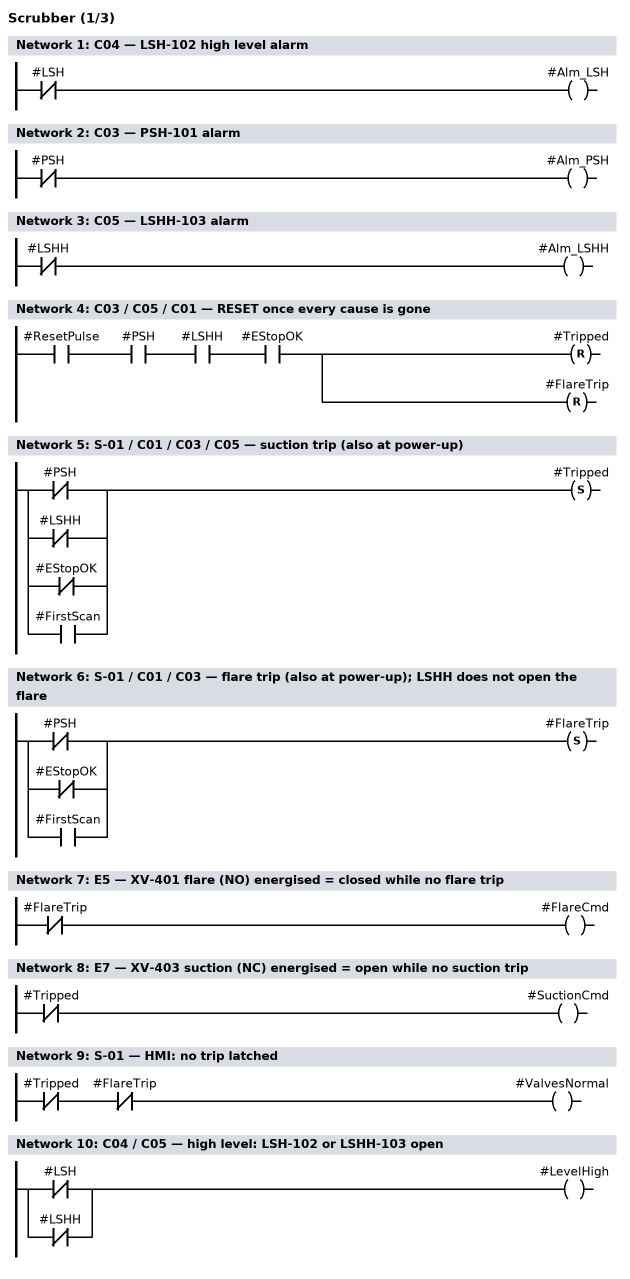
   RUNG wire#powerrail
      I_Contact( #LSH )
      Coil( #Alm_LSH )
   END_RUNG
   // the same network as SCL:
   #Alm_LSH := NOT #LSH;
END_REGION

REGION Network 2: C03 — PSH-101 alarm
   RUNG wire#powerrail
      I_Contact( #PSH )
      Coil( #Alm_PSH )
   END_RUNG
   // the same network as SCL:
   #Alm_PSH := NOT #PSH;
END_REGION

REGION Network 3: C05 — LSHH-103 alarm
   RUNG wire#powerrail
      I_Contact( #LSHH )
      Coil( #Alm_LSHH )
   END_RUNG
   // the same network as SCL:
   #Alm_LSHH := NOT #LSHH;
END_REGION

REGION Network 4: C03 / C05 / C01 — RESET once every cause is gone
   RUNG wire#powerrail
      Contact( #ResetPulse )
      Contact( #PSH )
      Contact( #LSHH )
      Contact( #EStopOK )
      wire#w1
      R_Coil( #Tripped )
   END_RUNG
   RUNG wire#w1
      R_Coil( #FlareTrip )
   END_RUNG
   // the same network as SCL:
   IF #ResetPulse AND #PSH AND #LSHH AND #EStopOK THEN
       #Tripped := FALSE;
       #FlareTrip := FALSE;
   END_IF;
END_REGION

REGION Network 5: S-01 / C01 / C03 / C05 — suction trip (also at power-up)
   RUNG wire#powerrail
      I_Contact( #PSH )
      wire#w1
      S_Coil( #Tripped )
   END_RUNG
   RUNG wire#powerrail
      I_Contact( #LSHH )
   END_RUNG wire#w1
   RUNG wire#powerrail
      I_Contact( #EStopOK )
   END_RUNG wire#w1
   RUNG wire#powerrail
      Contact( #FirstScan )
   END_RUNG wire#w1
   // the same network as SCL:
   IF NOT #PSH OR NOT #LSHH OR NOT #EStopOK OR #FirstScan THEN #Tripped := TRUE; END_IF;
END_REGION

REGION Network 6: S-01 / C01 / C03 — flare trip (also at power-up); LSHH does not open the flare
   RUNG wire#powerrail
      I_Contact( #PSH )
      wire#w1
      S_Coil( #FlareTrip )
   END_RUNG
   RUNG wire#powerrail
      I_Contact( #EStopOK )
   END_RUNG wire#w1
   RUNG wire#powerrail
      Contact( #FirstScan )
   END_RUNG wire#w1
   // the same network as SCL:
   IF NOT #PSH OR NOT #EStopOK OR #FirstScan THEN #FlareTrip := TRUE; END_IF;
END_REGION

REGION Network 7: E5 — XV-401 flare (NO) energised = closed while no flare trip
   RUNG wire#powerrail
      I_Contact( #FlareTrip )
      Coil( #FlareCmd )
   END_RUNG
   // the same network as SCL:
   #FlareCmd := NOT #FlareTrip;
END_REGION

REGION Network 8: E7 — XV-403 suction (NC) energised = open while no suction trip
   RUNG wire#powerrail
      I_Contact( #Tripped )
      Coil( #SuctionCmd )
   END_RUNG
   // the same network as SCL:
   #SuctionCmd := NOT #Tripped;
END_REGION

REGION Network 9: S-01 — HMI: no trip latched
   RUNG wire#powerrail
      I_Contact( #Tripped )
      I_Contact( #FlareTrip )
      Coil( #ValvesNormal )
   END_RUNG
   // the same network as SCL:
   #ValvesNormal := NOT #Tripped AND NOT #FlareTrip;
END_REGION

REGION Network 10: C04 / C05 — high level: LSH-102 or LSHH-103 open
   RUNG wire#powerrail
      I_Contact( #LSH )
      wire#w1
      Coil( #LevelHigh )
   END_RUNG
   RUNG wire#powerrail
      I_Contact( #LSHH )
   END_RUNG wire#w1
   // the same network as SCL:
   #LevelHigh := NOT #LSH OR NOT #LSHH;
END_REGION

REGION Network 11: C04 — drain demand after TDRN_ON of high level
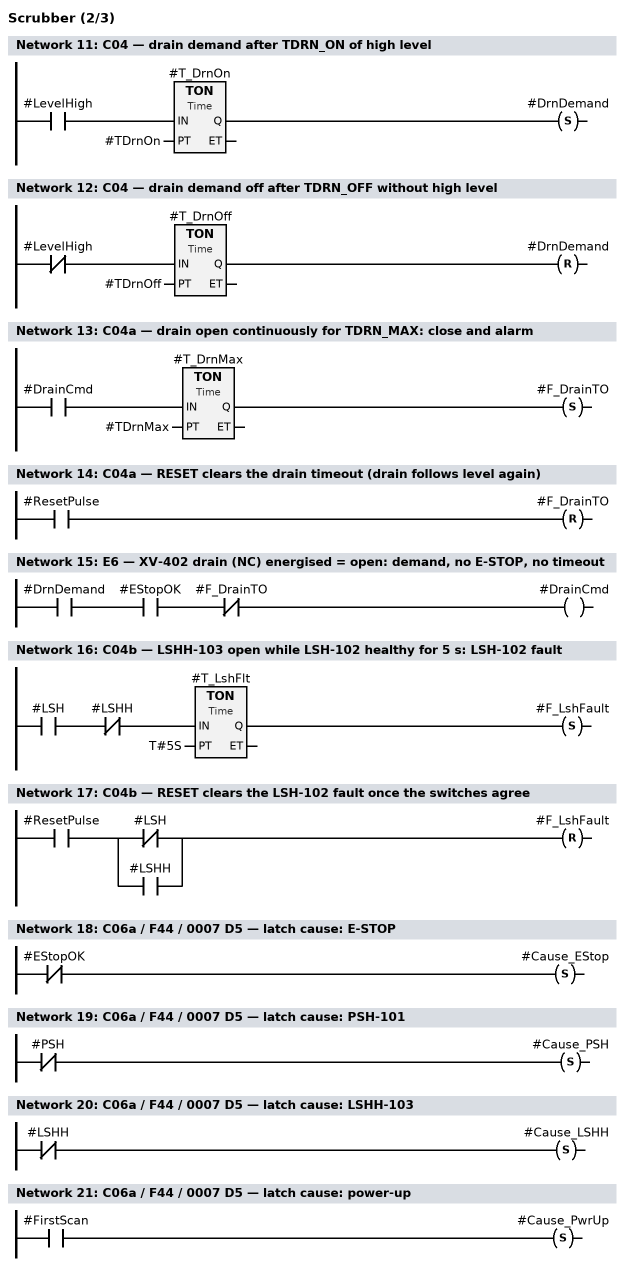
   RUNG wire#powerrail
      Contact( #LevelHigh )
      { S7_Templates := "time_type := Time" } #T_DrnOn.TON(pt := #TDrnOn, et =>)
      S_Coil( #DrnDemand )
   END_RUNG
   // the same network as SCL:
   #T_DrnOn(IN := #LevelHigh, PT := #TDrnOn);   // TON
   IF #T_DrnOn.Q THEN #DrnDemand := TRUE; END_IF;
END_REGION

REGION Network 12: C04 — drain demand off after TDRN_OFF without high level
   RUNG wire#powerrail
      I_Contact( #LevelHigh )
      { S7_Templates := "time_type := Time" } #T_DrnOff.TON(pt := #TDrnOff, et =>)
      R_Coil( #DrnDemand )
   END_RUNG
   // the same network as SCL:
   #T_DrnOff(IN := NOT #LevelHigh, PT := #TDrnOff);   // TON
   IF #T_DrnOff.Q THEN #DrnDemand := FALSE; END_IF;
END_REGION

REGION Network 13: C04a — drain open continuously for TDRN_MAX: close and alarm
   RUNG wire#powerrail
      Contact( #DrainCmd )
      { S7_Templates := "time_type := Time" } #T_DrnMax.TON(pt := #TDrnMax, et =>)
      S_Coil( #F_DrainTO )
   END_RUNG
   // the same network as SCL:
   #T_DrnMax(IN := #DrainCmd, PT := #TDrnMax);   // TON
   IF #T_DrnMax.Q THEN #F_DrainTO := TRUE; END_IF;
END_REGION

REGION Network 14: C04a — RESET clears the drain timeout (drain follows level again)
   RUNG wire#powerrail
      Contact( #ResetPulse )
      R_Coil( #F_DrainTO )
   END_RUNG
   // the same network as SCL:
   IF #ResetPulse THEN #F_DrainTO := FALSE; END_IF;
END_REGION

REGION Network 15: E6 — XV-402 drain (NC) energised = open: demand, no E-STOP, no timeout
   RUNG wire#powerrail
      Contact( #DrnDemand )
      Contact( #EStopOK )
      I_Contact( #F_DrainTO )
      Coil( #DrainCmd )
   END_RUNG
   // the same network as SCL:
   #DrainCmd := #DrnDemand AND #EStopOK AND NOT #F_DrainTO;
END_REGION

REGION Network 16: C04b — LSHH-103 open while LSH-102 healthy for 5 s: LSH-102 fault
   RUNG wire#powerrail
      Contact( #LSH )
      I_Contact( #LSHH )
      { S7_Templates := "time_type := Time" } #T_LshFlt.TON(pt := T#5S, et =>)
      S_Coil( #F_LshFault )
   END_RUNG
   // the same network as SCL:
   #T_LshFlt(IN := #LSH AND NOT #LSHH, PT := T#5S);   // TON
   IF #T_LshFlt.Q THEN #F_LshFault := TRUE; END_IF;
END_REGION

REGION Network 17: C04b — RESET clears the LSH-102 fault once the switches agree
   RUNG wire#powerrail
      Contact( #ResetPulse )
      wire#w1
      I_Contact( #LSH )
      wire#w2
      R_Coil( #F_LshFault )
   END_RUNG
   RUNG wire#w1
      Contact( #LSHH )
   END_RUNG wire#w2
   // the same network as SCL:
   IF #ResetPulse AND (NOT #LSH OR #LSHH) THEN #F_LshFault := FALSE; END_IF;
END_REGION

REGION Network 18: C06a / F44 / 0007 D5 — latch cause: E-STOP
   RUNG wire#powerrail
      I_Contact( #EStopOK )
      S_Coil( #Cause_EStop )
   END_RUNG
   // the same network as SCL:
   IF NOT #EStopOK THEN #Cause_EStop := TRUE; END_IF;
END_REGION

REGION Network 19: C06a / F44 / 0007 D5 — latch cause: PSH-101
   RUNG wire#powerrail
      I_Contact( #PSH )
      S_Coil( #Cause_PSH )
   END_RUNG
   // the same network as SCL:
   IF NOT #PSH THEN #Cause_PSH := TRUE; END_IF;
END_REGION

REGION Network 20: C06a / F44 / 0007 D5 — latch cause: LSHH-103
   RUNG wire#powerrail
      I_Contact( #LSHH )
      S_Coil( #Cause_LSHH )
   END_RUNG
   // the same network as SCL:
   IF NOT #LSHH THEN #Cause_LSHH := TRUE; END_IF;
END_REGION

REGION Network 21: C06a / F44 / 0007 D5 — latch cause: power-up
   RUNG wire#powerrail
      Contact( #FirstScan )
      S_Coil( #Cause_PwrUp )
   END_RUNG
   // the same network as SCL:
   IF #FirstScan THEN #Cause_PwrUp := TRUE; END_IF;
END_REGION

REGION Network 22: C06a / F44 / 0007 D5 — first-out 1: E-STOP (only if none)
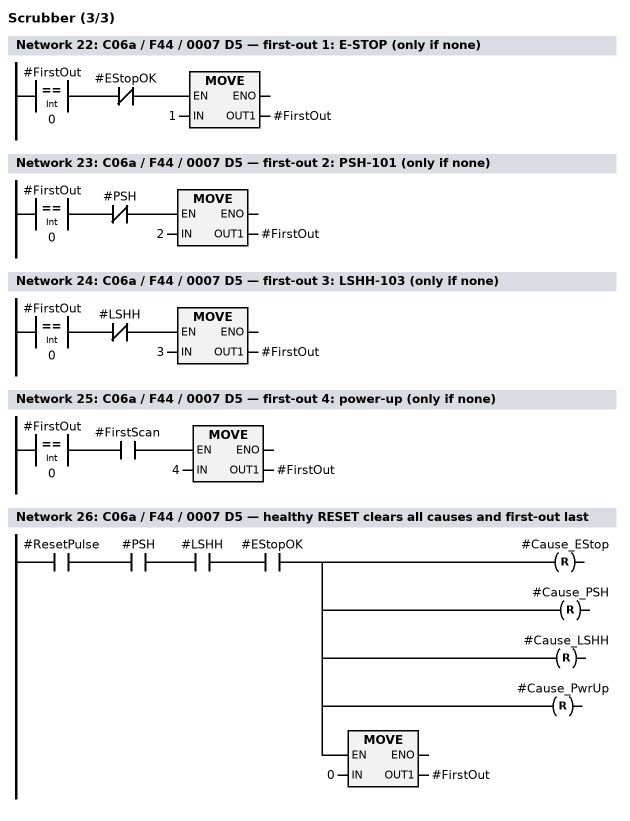
   RUNG wire#powerrail
      { S7_Templates := "SrcType := Int" } EQ_Contact(in1 := #FirstOut, in2 := 0)
      I_Contact( #EStopOK )
      { S7_GenerateENO := "TRUE" } Move(in := 1, out1 => #FirstOut)
   END_RUNG
   // the same network as SCL:
   IF (#FirstOut = 0) AND NOT #EStopOK THEN #FirstOut := 1; END_IF;
END_REGION

REGION Network 23: C06a / F44 / 0007 D5 — first-out 2: PSH-101 (only if none)
   RUNG wire#powerrail
      { S7_Templates := "SrcType := Int" } EQ_Contact(in1 := #FirstOut, in2 := 0)
      I_Contact( #PSH )
      { S7_GenerateENO := "TRUE" } Move(in := 2, out1 => #FirstOut)
   END_RUNG
   // the same network as SCL:
   IF (#FirstOut = 0) AND NOT #PSH THEN #FirstOut := 2; END_IF;
END_REGION

REGION Network 24: C06a / F44 / 0007 D5 — first-out 3: LSHH-103 (only if none)
   RUNG wire#powerrail
      { S7_Templates := "SrcType := Int" } EQ_Contact(in1 := #FirstOut, in2 := 0)
      I_Contact( #LSHH )
      { S7_GenerateENO := "TRUE" } Move(in := 3, out1 => #FirstOut)
   END_RUNG
   // the same network as SCL:
   IF (#FirstOut = 0) AND NOT #LSHH THEN #FirstOut := 3; END_IF;
END_REGION

REGION Network 25: C06a / F44 / 0007 D5 — first-out 4: power-up (only if none)
   RUNG wire#powerrail
      { S7_Templates := "SrcType := Int" } EQ_Contact(in1 := #FirstOut, in2 := 0)
      Contact( #FirstScan )
      { S7_GenerateENO := "TRUE" } Move(in := 4, out1 => #FirstOut)
   END_RUNG
   // the same network as SCL:
   IF (#FirstOut = 0) AND #FirstScan THEN #FirstOut := 4; END_IF;
END_REGION

REGION Network 26: C06a / F44 / 0007 D5 — healthy RESET clears all causes and first-out last
   RUNG wire#powerrail
      Contact( #ResetPulse )
      Contact( #PSH )
      Contact( #LSHH )
      Contact( #EStopOK )
      wire#w1
      R_Coil( #Cause_EStop )
   END_RUNG
   RUNG wire#w1
      R_Coil( #Cause_PSH )
   END_RUNG
   RUNG wire#w1
      R_Coil( #Cause_LSHH )
   END_RUNG
   RUNG wire#w1
      R_Coil( #Cause_PwrUp )
   END_RUNG
   RUNG wire#w1
      { S7_GenerateENO := "TRUE" } Move(in := 0, out1 => #FirstOut)
   END_RUNG
   // the same network as SCL:
   IF #ResetPulse AND #PSH AND #LSHH AND #EStopOK THEN
       #Cause_EStop := FALSE;
       #Cause_PSH := FALSE;
       #Cause_LSHH := FALSE;
       #Cause_PwrUp := FALSE;
       #FirstOut := 0;
   END_IF;
END_REGION
END_FUNCTION_BLOCK

FUNCTION_BLOCK "Burner"   // FB1, LAD
TITLE = Burner
{ S7_Optimized_Access := 'TRUE' }
VERSION : 0.1
// One burner, docs/التشغيل.md §2 and decisions/0006
// stored: AutoNumber false, IsIECCheckEnabled false, MemoryReserve 100, SetENOAutomatically False
   VAR_INPUT
      Auto : Bool;   // AUTO/MAN selector, 1 = AUTO
      StartPB : Bool;   // START push button (NO)
      StopOK : Bool;   // STOP push button (NC): 1 = released
      LevelOK : Bool;   // Tank LSL reached (C07a)
      RunFb : Bool;   // Burner RUN feedback
      Lockout : Bool;   // Burner lockout signal (C07e)
      Fuel : Bool;   // Fuel mode (BR02 Rfuel2, R-12); FALSE for BR01
      TeA : Int;   // Thermocouple A raw, 0.1 degC
      TeB : Int;   // Thermocouple B raw, 0.1 degC
      Use24h : Bool;   // 24 h forced stop enabled (C07h, BR01 only)
      EStopOK : Bool;   // Sys.EStopOK
      ResetPulse : Bool;   // Sys.ResetPulse
      FirstScan : Bool;   // Sys.FirstScan
      SP : Int;   // Par.SP_V
      HYST : Int;   // Par.HYST_V
      STG : Int;   // Par.STG_V
      TStart : Time;   // Par.TStart_V
   END_VAR
   VAR_OUTPUT
      HeatReq : Bool;   // Heat request TL / L (E1 / E3)
      Stage2 : Bool;   // 2nd stage TR / T2 (E2 / E4)
      State : Int;   // 0 IDLE, 1 STARTING, 2 RUNNING, 3 FAULT
      Enabled : Bool;   // START given and not taken back (B-01)
      Tmax : Int;   // Higher of the two thermocouples, 0.1 degC
      F_EStop : Bool;   // Fault C01
      F_TC : Bool;   // Fault C0xd thermocouple
      F_Lockout : Bool;   // Fault C0xe lockout
      F_NoStart : Bool;   // Fault C0xf failed to start
      F_RunLost : Bool;   // Fault C0xg stopped by itself
      F_RunWrong : Bool;   // Fault R-09 RUN without request
      ParPending : Bool;   // R-11 / D6 / 0007: a validated entry differs from its active copy
   END_VAR
   VAR
      StartEdge : Bool;
      StartMem : Bool;
      AutoChg : Bool;
      AutoMem : Bool;
      FuelChg : Bool;
      FuelMem : Bool;
      TcOkA : Bool;
      TcOkB : Bool;
      TcOk : Bool;
      TcBad : Bool;
      Demand : Bool;
      HeatNeed : Bool;
      Ready : Bool;
      Active : Bool;
      Pause24 : Bool;
      RunWrong : Bool;
      NoStart : Bool;
      PwrUpDone : Bool;
      TcSlow : Bool;
      SP_Act : Int;
      HYST_Act : Int;
      STG_Act : Int;
      TStart_Act : Time;
      TOn : Int;
      TStg : Int;
      TStgOff : Int;
      T_PwrUp : TON_TIME;
      T_TcBad : TON_TIME;
      T_24h : TON_TIME;
      T_Pause : TON_TIME;
      T_RunOff : TON_TIME;
      T_Start : TON_TIME;
   END_VAR
   VAR_TEMP   // added for the SCL form of the ladder/FBD networks
      _w1 : Bool;
   END_VAR
BEGIN

REGION Network 1: R-05 — START edge: not on first scan, only after seen released, STOP wins
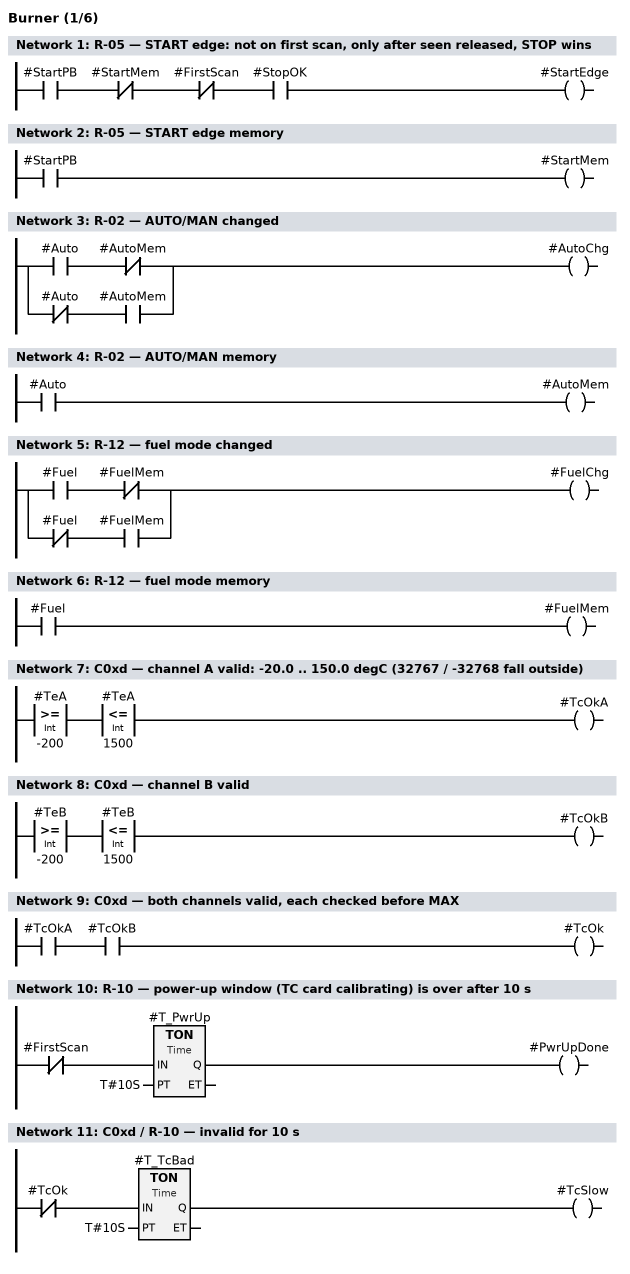
   RUNG wire#powerrail
      Contact( #StartPB )
      I_Contact( #StartMem )
      I_Contact( #FirstScan )
      Contact( #StopOK )
      Coil( #StartEdge )
   END_RUNG
   // the same network as SCL:
   #StartEdge := #StartPB AND NOT #StartMem AND NOT #FirstScan AND #StopOK;
END_REGION

REGION Network 2: R-05 — START edge memory
   RUNG wire#powerrail
      Contact( #StartPB )
      Coil( #StartMem )
   END_RUNG
   // the same network as SCL:
   #StartMem := #StartPB;
END_REGION

REGION Network 3: R-02 — AUTO/MAN changed
   RUNG wire#powerrail
      Contact( #Auto )
      I_Contact( #AutoMem )
      wire#w1
      Coil( #AutoChg )
   END_RUNG
   RUNG wire#powerrail
      I_Contact( #Auto )
      Contact( #AutoMem )
   END_RUNG wire#w1
   // the same network as SCL:
   #AutoChg := (#Auto AND NOT #AutoMem) OR (NOT #Auto AND #AutoMem);
END_REGION

REGION Network 4: R-02 — AUTO/MAN memory
   RUNG wire#powerrail
      Contact( #Auto )
      Coil( #AutoMem )
   END_RUNG
   // the same network as SCL:
   #AutoMem := #Auto;
END_REGION

REGION Network 5: R-12 — fuel mode changed
   RUNG wire#powerrail
      Contact( #Fuel )
      I_Contact( #FuelMem )
      wire#w1
      Coil( #FuelChg )
   END_RUNG
   RUNG wire#powerrail
      I_Contact( #Fuel )
      Contact( #FuelMem )
   END_RUNG wire#w1
   // the same network as SCL:
   #FuelChg := (#Fuel AND NOT #FuelMem) OR (NOT #Fuel AND #FuelMem);
END_REGION

REGION Network 6: R-12 — fuel mode memory
   RUNG wire#powerrail
      Contact( #Fuel )
      Coil( #FuelMem )
   END_RUNG
   // the same network as SCL:
   #FuelMem := #Fuel;
END_REGION

REGION Network 7: C0xd — channel A valid: -20.0 .. 150.0 degC (32767 / -32768 fall outside)
   RUNG wire#powerrail
      { S7_Templates := "SrcType := Int" } GE_Contact(in1 := #TeA, in2 := -200)
      { S7_Templates := "SrcType := Int" } LE_Contact(in1 := #TeA, in2 := 1500)
      Coil( #TcOkA )
   END_RUNG
   // the same network as SCL:
   #TcOkA := (#TeA >= (-200)) AND (#TeA <= 1500);
END_REGION

REGION Network 8: C0xd — channel B valid
   RUNG wire#powerrail
      { S7_Templates := "SrcType := Int" } GE_Contact(in1 := #TeB, in2 := -200)
      { S7_Templates := "SrcType := Int" } LE_Contact(in1 := #TeB, in2 := 1500)
      Coil( #TcOkB )
   END_RUNG
   // the same network as SCL:
   #TcOkB := (#TeB >= (-200)) AND (#TeB <= 1500);
END_REGION

REGION Network 9: C0xd — both channels valid, each checked before MAX
   RUNG wire#powerrail
      Contact( #TcOkA )
      Contact( #TcOkB )
      Coil( #TcOk )
   END_RUNG
   // the same network as SCL:
   #TcOk := #TcOkA AND #TcOkB;
END_REGION

REGION Network 10: R-10 — power-up window (TC card calibrating) is over after 10 s
   RUNG wire#powerrail
      I_Contact( #FirstScan )
      { S7_Templates := "time_type := Time" } #T_PwrUp.TON(pt := T#10S, et =>)
      Coil( #PwrUpDone )
   END_RUNG
   // the same network as SCL:
   #T_PwrUp(IN := NOT #FirstScan, PT := T#10S);   // TON
   #PwrUpDone := #T_PwrUp.Q;
END_REGION

REGION Network 11: C0xd / R-10 — invalid for 10 s
   RUNG wire#powerrail
      I_Contact( #TcOk )
      { S7_Templates := "time_type := Time" } #T_TcBad.TON(pt := T#10S, et =>)
      Coil( #TcSlow )
   END_RUNG
   // the same network as SCL:
   #T_TcBad(IN := NOT #TcOk, PT := T#10S);   // TON
   #TcSlow := #T_TcBad.Q;
END_REGION

REGION Network 12: C0xd / R-10 — invalid = fault: at once, or after 10 s right after power-up
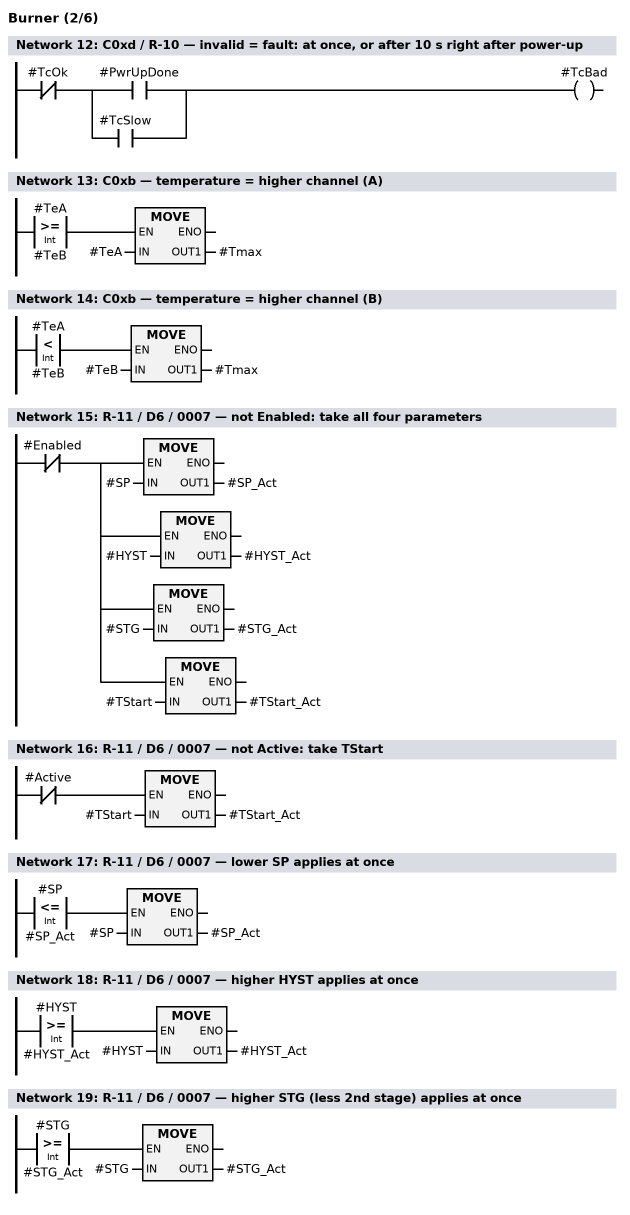
   RUNG wire#powerrail
      I_Contact( #TcOk )
      wire#w1
      Contact( #PwrUpDone )
      wire#w2
      Coil( #TcBad )
   END_RUNG
   RUNG wire#w1
      Contact( #TcSlow )
   END_RUNG wire#w2
   // the same network as SCL:
   #TcBad := NOT #TcOk AND (#PwrUpDone OR #TcSlow);
END_REGION

REGION Network 13: C0xb — temperature = higher channel (A)
   RUNG wire#powerrail
      { S7_Templates := "SrcType := Int" } GE_Contact(in1 := #TeA, in2 := #TeB)
      { S7_GenerateENO := "TRUE" } Move(in := #TeA, out1 => #Tmax)
   END_RUNG
   // the same network as SCL:
   IF #TeA >= #TeB THEN #Tmax := #TeA; END_IF;
END_REGION

REGION Network 14: C0xb — temperature = higher channel (B)
   RUNG wire#powerrail
      { S7_Templates := "SrcType := Int" } LT_Contact(in1 := #TeA, in2 := #TeB)
      { S7_GenerateENO := "TRUE" } Move(in := #TeB, out1 => #Tmax)
   END_RUNG
   // the same network as SCL:
   IF #TeA < #TeB THEN #Tmax := #TeB; END_IF;
END_REGION

REGION Network 15: R-11 / D6 / 0007 — not Enabled: take all four parameters
   RUNG wire#powerrail
      I_Contact( #Enabled )
      wire#w1
      { S7_GenerateENO := "TRUE" } Move(in := #SP, out1 => #SP_Act)
   END_RUNG
   RUNG wire#w1
      { S7_GenerateENO := "TRUE" } Move(in := #HYST, out1 => #HYST_Act)
   END_RUNG
   RUNG wire#w1
      { S7_GenerateENO := "TRUE" } Move(in := #STG, out1 => #STG_Act)
   END_RUNG
   RUNG wire#w1
      { S7_GenerateENO := "TRUE" } Move(in := #TStart, out1 => #TStart_Act)
   END_RUNG
   // the same network as SCL:
   IF NOT #Enabled THEN
       #SP_Act := #SP;
       #HYST_Act := #HYST;
       #STG_Act := #STG;
       #TStart_Act := #TStart;
   END_IF;
END_REGION

REGION Network 16: R-11 / D6 / 0007 — not Active: take TStart
   RUNG wire#powerrail
      I_Contact( #Active )
      { S7_GenerateENO := "TRUE" } Move(in := #TStart, out1 => #TStart_Act)
   END_RUNG
   // the same network as SCL:
   IF NOT #Active THEN #TStart_Act := #TStart; END_IF;
END_REGION

REGION Network 17: R-11 / D6 / 0007 — lower SP applies at once
   RUNG wire#powerrail
      { S7_Templates := "SrcType := Int" } LE_Contact(in1 := #SP, in2 := #SP_Act)
      { S7_GenerateENO := "TRUE" } Move(in := #SP, out1 => #SP_Act)
   END_RUNG
   // the same network as SCL:
   IF #SP <= #SP_Act THEN #SP_Act := #SP; END_IF;
END_REGION

REGION Network 18: R-11 / D6 / 0007 — higher HYST applies at once
   RUNG wire#powerrail
      { S7_Templates := "SrcType := Int" } GE_Contact(in1 := #HYST, in2 := #HYST_Act)
      { S7_GenerateENO := "TRUE" } Move(in := #HYST, out1 => #HYST_Act)
   END_RUNG
   // the same network as SCL:
   IF #HYST >= #HYST_Act THEN #HYST_Act := #HYST; END_IF;
END_REGION

REGION Network 19: R-11 / D6 / 0007 — higher STG (less 2nd stage) applies at once
   RUNG wire#powerrail
      { S7_Templates := "SrcType := Int" } GE_Contact(in1 := #STG, in2 := #STG_Act)
      { S7_GenerateENO := "TRUE" } Move(in := #STG, out1 => #STG_Act)
   END_RUNG
   // the same network as SCL:
   IF #STG >= #STG_Act THEN #STG_Act := #STG; END_IF;
END_REGION

REGION Network 20: R-11 / D6 / 0007 — pending while any entry differs from its active copy
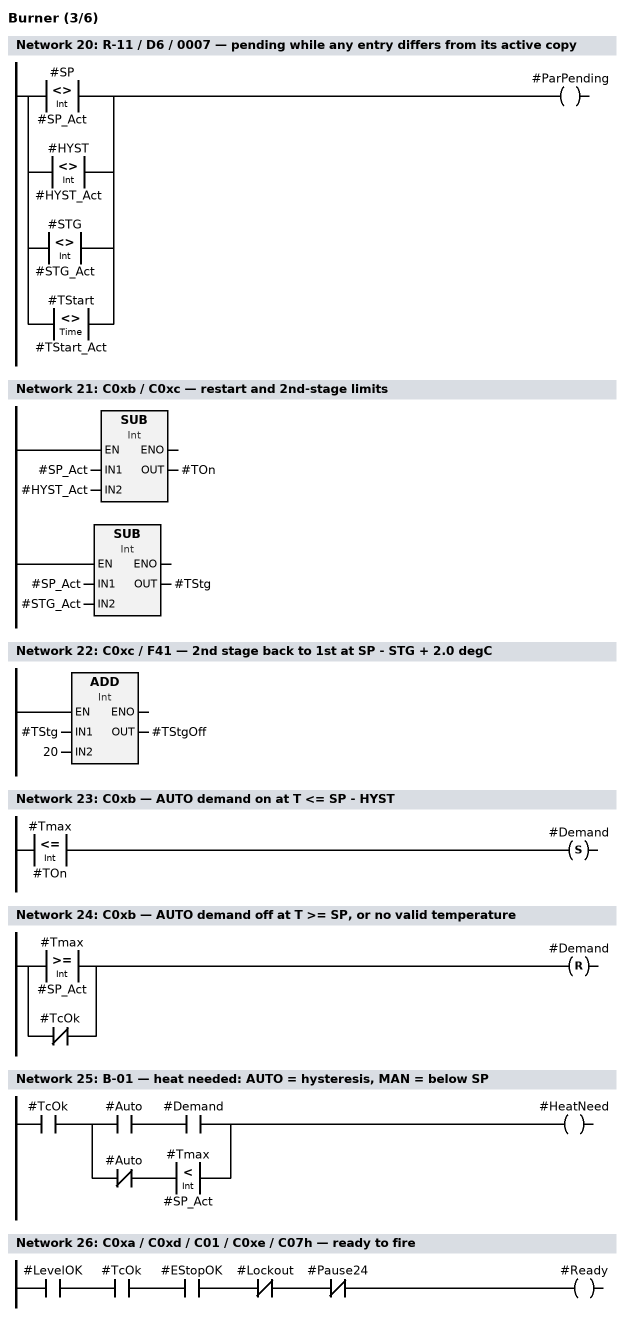
   RUNG wire#powerrail
      { S7_Templates := "SrcType := Int" } NE_Contact(in1 := #SP, in2 := #SP_Act)
      wire#w1
      Coil( #ParPending )
   END_RUNG
   RUNG wire#powerrail
      { S7_Templates := "SrcType := Int" } NE_Contact(in1 := #HYST, in2 := #HYST_Act)
   END_RUNG wire#w1
   RUNG wire#powerrail
      { S7_Templates := "SrcType := Int" } NE_Contact(in1 := #STG, in2 := #STG_Act)
   END_RUNG wire#w1
   RUNG wire#powerrail
      { S7_Templates := "SrcType := Time" } NE_Contact(in1 := #TStart, in2 := #TStart_Act)
   END_RUNG wire#w1
   // the same network as SCL:
   #ParPending := (#SP <> #SP_Act) OR (#HYST <> #HYST_Act) OR (#STG <> #STG_Act) OR (#TStart <> #TStart_Act);
END_REGION

REGION Network 21: C0xb / C0xc — restart and 2nd-stage limits
   RUNG wire#powerrail
      { S7_Templates := "SrcType := Int"; S7_GenerateENO := "TRUE" } Sub(in1 := #SP_Act, in2 := #HYST_Act, out => #TOn)
   END_RUNG
   RUNG wire#powerrail
      { S7_Templates := "SrcType := Int"; S7_GenerateENO := "TRUE" } Sub(in1 := #SP_Act, in2 := #STG_Act, out => #TStg)
   END_RUNG
   // the same network as SCL:
   #TOn := #SP_Act - #HYST_Act;
   #TStg := #SP_Act - #STG_Act;
END_REGION

REGION Network 22: C0xc / F41 — 2nd stage back to 1st at SP - STG + 2.0 degC
   RUNG wire#powerrail
      { S7_Templates := "SrcType := Int"; S7_GenerateENO := "TRUE" } Add(in1 := #TStg, in2 := 20, out => #TStgOff)
   END_RUNG
   // the same network as SCL:
   #TStgOff := #TStg + 20;
END_REGION

REGION Network 23: C0xb — AUTO demand on at T <= SP - HYST
   RUNG wire#powerrail
      { S7_Templates := "SrcType := Int" } LE_Contact(in1 := #Tmax, in2 := #TOn)
      S_Coil( #Demand )
   END_RUNG
   // the same network as SCL:
   IF #Tmax <= #TOn THEN #Demand := TRUE; END_IF;
END_REGION

REGION Network 24: C0xb — AUTO demand off at T >= SP, or no valid temperature
   RUNG wire#powerrail
      { S7_Templates := "SrcType := Int" } GE_Contact(in1 := #Tmax, in2 := #SP_Act)
      wire#w1
      R_Coil( #Demand )
   END_RUNG
   RUNG wire#powerrail
      I_Contact( #TcOk )
   END_RUNG wire#w1
   // the same network as SCL:
   IF (#Tmax >= #SP_Act) OR NOT #TcOk THEN #Demand := FALSE; END_IF;
END_REGION

REGION Network 25: B-01 — heat needed: AUTO = hysteresis, MAN = below SP
   RUNG wire#powerrail
      Contact( #TcOk )
      wire#w1
      Contact( #Auto )
      Contact( #Demand )
      wire#w2
      Coil( #HeatNeed )
   END_RUNG
   RUNG wire#w1
      I_Contact( #Auto )
      { S7_Templates := "SrcType := Int" } LT_Contact(in1 := #Tmax, in2 := #SP_Act)
   END_RUNG wire#w2
   // the same network as SCL:
   #HeatNeed := #TcOk AND ((#Auto AND #Demand) OR (NOT #Auto AND (#Tmax < #SP_Act)));
END_REGION

REGION Network 26: C0xa / C0xd / C01 / C0xe / C07h — ready to fire
   RUNG wire#powerrail
      Contact( #LevelOK )
      Contact( #TcOk )
      Contact( #EStopOK )
      I_Contact( #Lockout )
      I_Contact( #Pause24 )
      Coil( #Ready )
   END_RUNG
   // the same network as SCL:
   #Ready := #LevelOK AND #TcOk AND #EStopOK AND NOT #Lockout AND NOT #Pause24;
END_REGION

REGION Network 27: C07h / R-08 — 24 h of continuous request: forced stop
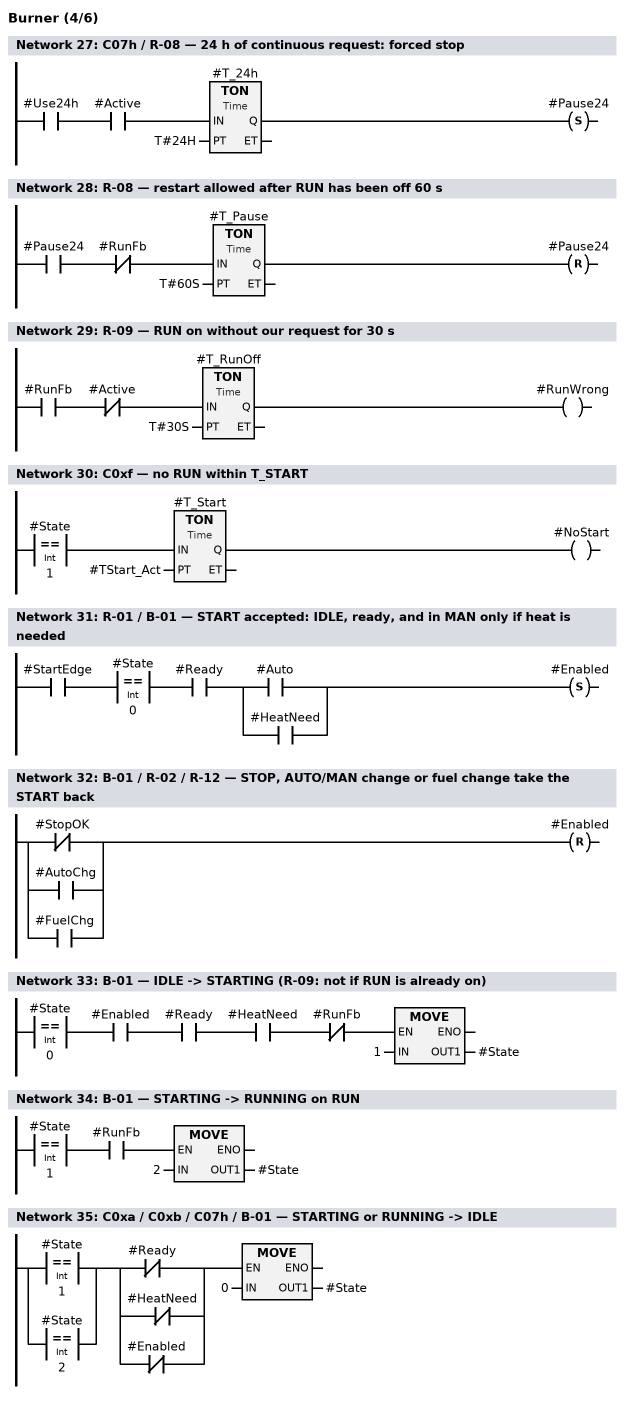
   RUNG wire#powerrail
      Contact( #Use24h )
      Contact( #Active )
      { S7_Templates := "time_type := Time" } #T_24h.TON(pt := T#24H, et =>)
      S_Coil( #Pause24 )
   END_RUNG
   // the same network as SCL:
   #T_24h(IN := #Use24h AND #Active, PT := T#24H);   // TON
   IF #T_24h.Q THEN #Pause24 := TRUE; END_IF;
END_REGION

REGION Network 28: R-08 — restart allowed after RUN has been off 60 s
   RUNG wire#powerrail
      Contact( #Pause24 )
      I_Contact( #RunFb )
      { S7_Templates := "time_type := Time" } #T_Pause.TON(pt := T#60S, et =>)
      R_Coil( #Pause24 )
   END_RUNG
   // the same network as SCL:
   #T_Pause(IN := #Pause24 AND NOT #RunFb, PT := T#60S);   // TON
   IF #T_Pause.Q THEN #Pause24 := FALSE; END_IF;
END_REGION

REGION Network 29: R-09 — RUN on without our request for 30 s
   RUNG wire#powerrail
      Contact( #RunFb )
      I_Contact( #Active )
      { S7_Templates := "time_type := Time" } #T_RunOff.TON(pt := T#30S, et =>)
      Coil( #RunWrong )
   END_RUNG
   // the same network as SCL:
   #T_RunOff(IN := #RunFb AND NOT #Active, PT := T#30S);   // TON
   #RunWrong := #T_RunOff.Q;
END_REGION

REGION Network 30: C0xf — no RUN within T_START
   RUNG wire#powerrail
      { S7_Templates := "SrcType := Int" } EQ_Contact(in1 := #State, in2 := 1)
      { S7_Templates := "time_type := Time" } #T_Start.TON(pt := #TStart_Act, et =>)
      Coil( #NoStart )
   END_RUNG
   // the same network as SCL:
   #T_Start(IN := #State = 1, PT := #TStart_Act);   // TON
   #NoStart := #T_Start.Q;
END_REGION

REGION Network 31: R-01 / B-01 — START accepted: IDLE, ready, and in MAN only if heat is needed
   RUNG wire#powerrail
      Contact( #StartEdge )
      { S7_Templates := "SrcType := Int" } EQ_Contact(in1 := #State, in2 := 0)
      Contact( #Ready )
      wire#w1
      Contact( #Auto )
      wire#w2
      S_Coil( #Enabled )
   END_RUNG
   RUNG wire#w1
      Contact( #HeatNeed )
   END_RUNG wire#w2
   // the same network as SCL:
   IF #StartEdge AND (#State = 0) AND #Ready AND (#Auto OR #HeatNeed) THEN #Enabled := TRUE; END_IF;
END_REGION

REGION Network 32: B-01 / R-02 / R-12 — STOP, AUTO/MAN change or fuel change take the START back
   RUNG wire#powerrail
      I_Contact( #StopOK )
      wire#w1
      R_Coil( #Enabled )
   END_RUNG
   RUNG wire#powerrail
      Contact( #AutoChg )
   END_RUNG wire#w1
   RUNG wire#powerrail
      Contact( #FuelChg )
   END_RUNG wire#w1
   // the same network as SCL:
   IF NOT #StopOK OR #AutoChg OR #FuelChg THEN #Enabled := FALSE; END_IF;
END_REGION

REGION Network 33: B-01 — IDLE -> STARTING (R-09: not if RUN is already on)
   RUNG wire#powerrail
      { S7_Templates := "SrcType := Int" } EQ_Contact(in1 := #State, in2 := 0)
      Contact( #Enabled )
      Contact( #Ready )
      Contact( #HeatNeed )
      I_Contact( #RunFb )
      { S7_GenerateENO := "TRUE" } Move(in := 1, out1 => #State)
   END_RUNG
   // the same network as SCL:
   IF (#State = 0) AND #Enabled AND #Ready AND #HeatNeed AND NOT #RunFb THEN #State := 1; END_IF;
END_REGION

REGION Network 34: B-01 — STARTING -> RUNNING on RUN
   RUNG wire#powerrail
      { S7_Templates := "SrcType := Int" } EQ_Contact(in1 := #State, in2 := 1)
      Contact( #RunFb )
      { S7_GenerateENO := "TRUE" } Move(in := 2, out1 => #State)
   END_RUNG
   // the same network as SCL:
   IF (#State = 1) AND #RunFb THEN #State := 2; END_IF;
END_REGION

REGION Network 35: C0xa / C0xb / C07h / B-01 — STARTING or RUNNING -> IDLE
   RUNG wire#powerrail
      { S7_Templates := "SrcType := Int" } EQ_Contact(in1 := #State, in2 := 1)
      wire#w1
      I_Contact( #Ready )
      wire#w2
      { S7_GenerateENO := "TRUE" } Move(in := 0, out1 => #State)
   END_RUNG
   RUNG wire#powerrail
      { S7_Templates := "SrcType := Int" } EQ_Contact(in1 := #State, in2 := 2)
   END_RUNG wire#w1
   RUNG wire#w1
      I_Contact( #HeatNeed )
   END_RUNG wire#w2
   RUNG wire#w1
      I_Contact( #Enabled )
   END_RUNG wire#w2
   // the same network as SCL:
   IF ((#State = 1) OR (#State = 2)) AND (NOT #Ready OR NOT #HeatNeed OR NOT #Enabled) THEN
       #State := 0;
   END_IF;
END_REGION

REGION Network 36: R-03 — MAN: one cycle; any stop needs a new START
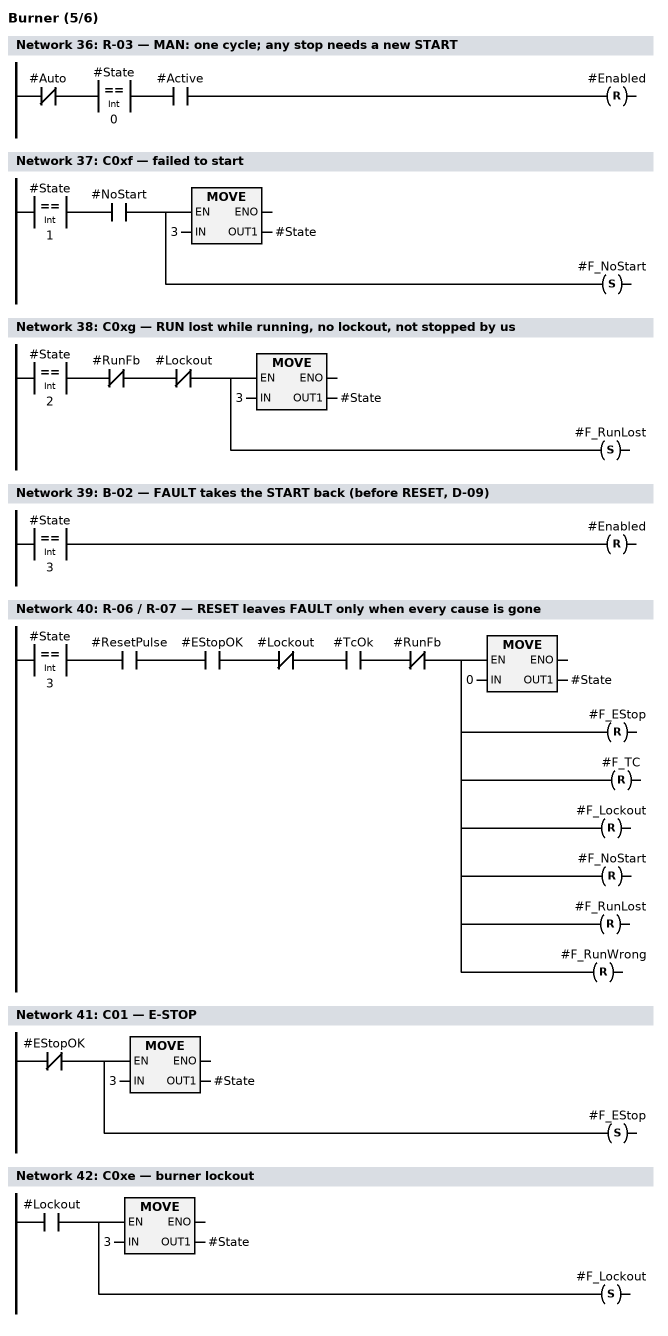
   RUNG wire#powerrail
      I_Contact( #Auto )
      { S7_Templates := "SrcType := Int" } EQ_Contact(in1 := #State, in2 := 0)
      Contact( #Active )
      R_Coil( #Enabled )
   END_RUNG
   // the same network as SCL:
   IF NOT #Auto AND (#State = 0) AND #Active THEN #Enabled := FALSE; END_IF;
END_REGION

REGION Network 37: C0xf — failed to start
   RUNG wire#powerrail
      { S7_Templates := "SrcType := Int" } EQ_Contact(in1 := #State, in2 := 1)
      Contact( #NoStart )
      wire#w1
      { S7_GenerateENO := "TRUE" } Move(in := 3, out1 => #State)
   END_RUNG
   RUNG wire#w1
      S_Coil( #F_NoStart )
   END_RUNG
   // the same network as SCL:
   #_w1 := (#State = 1) AND #NoStart;
   IF #_w1 THEN
       #State := 3;
       #F_NoStart := TRUE;
   END_IF;
END_REGION

REGION Network 38: C0xg — RUN lost while running, no lockout, not stopped by us
   RUNG wire#powerrail
      { S7_Templates := "SrcType := Int" } EQ_Contact(in1 := #State, in2 := 2)
      I_Contact( #RunFb )
      I_Contact( #Lockout )
      wire#w1
      { S7_GenerateENO := "TRUE" } Move(in := 3, out1 => #State)
   END_RUNG
   RUNG wire#w1
      S_Coil( #F_RunLost )
   END_RUNG
   // the same network as SCL:
   #_w1 := (#State = 2) AND NOT #RunFb AND NOT #Lockout;
   IF #_w1 THEN
       #State := 3;
       #F_RunLost := TRUE;
   END_IF;
END_REGION

REGION Network 39: B-02 — FAULT takes the START back (before RESET, D-09)
   RUNG wire#powerrail
      { S7_Templates := "SrcType := Int" } EQ_Contact(in1 := #State, in2 := 3)
      R_Coil( #Enabled )
   END_RUNG
   // the same network as SCL:
   IF #State = 3 THEN #Enabled := FALSE; END_IF;
END_REGION

REGION Network 40: R-06 / R-07 — RESET leaves FAULT only when every cause is gone
   RUNG wire#powerrail
      { S7_Templates := "SrcType := Int" } EQ_Contact(in1 := #State, in2 := 3)
      Contact( #ResetPulse )
      Contact( #EStopOK )
      I_Contact( #Lockout )
      Contact( #TcOk )
      I_Contact( #RunFb )
      wire#w1
      { S7_GenerateENO := "TRUE" } Move(in := 0, out1 => #State)
   END_RUNG
   RUNG wire#w1
      R_Coil( #F_EStop )
   END_RUNG
   RUNG wire#w1
      R_Coil( #F_TC )
   END_RUNG
   RUNG wire#w1
      R_Coil( #F_Lockout )
   END_RUNG
   RUNG wire#w1
      R_Coil( #F_NoStart )
   END_RUNG
   RUNG wire#w1
      R_Coil( #F_RunLost )
   END_RUNG
   RUNG wire#w1
      R_Coil( #F_RunWrong )
   END_RUNG
   // the same network as SCL:
   #_w1 := (#State = 3) AND #ResetPulse AND #EStopOK AND NOT #Lockout AND #TcOk AND NOT #RunFb;
   IF #_w1 THEN
       #State := 0;
       #F_EStop := FALSE;
       #F_TC := FALSE;
       #F_Lockout := FALSE;
       #F_NoStart := FALSE;
       #F_RunLost := FALSE;
       #F_RunWrong := FALSE;
   END_IF;
END_REGION

REGION Network 41: C01 — E-STOP
   RUNG wire#powerrail
      I_Contact( #EStopOK )
      wire#w1
      { S7_GenerateENO := "TRUE" } Move(in := 3, out1 => #State)
   END_RUNG
   RUNG wire#w1
      S_Coil( #F_EStop )
   END_RUNG
   // the same network as SCL:
   IF NOT #EStopOK THEN
       #State := 3;
       #F_EStop := TRUE;
   END_IF;
END_REGION

REGION Network 42: C0xe — burner lockout
   RUNG wire#powerrail
      Contact( #Lockout )
      wire#w1
      { S7_GenerateENO := "TRUE" } Move(in := 3, out1 => #State)
   END_RUNG
   RUNG wire#w1
      S_Coil( #F_Lockout )
   END_RUNG
   // the same network as SCL:
   IF #Lockout THEN
       #State := 3;
       #F_Lockout := TRUE;
   END_IF;
END_REGION

REGION Network 43: C0xd — thermocouple fault
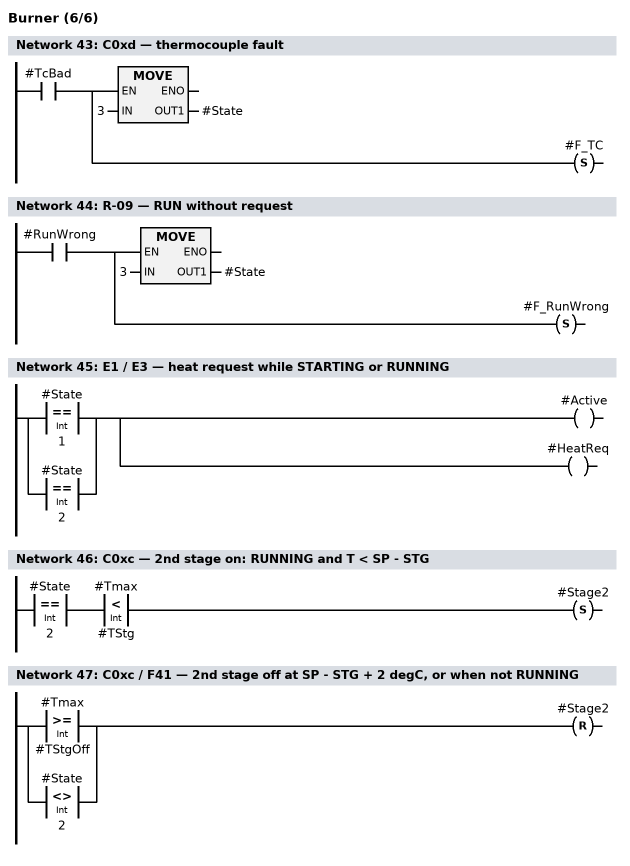
   RUNG wire#powerrail
      Contact( #TcBad )
      wire#w1
      { S7_GenerateENO := "TRUE" } Move(in := 3, out1 => #State)
   END_RUNG
   RUNG wire#w1
      S_Coil( #F_TC )
   END_RUNG
   // the same network as SCL:
   IF #TcBad THEN
       #State := 3;
       #F_TC := TRUE;
   END_IF;
END_REGION

REGION Network 44: R-09 — RUN without request
   RUNG wire#powerrail
      Contact( #RunWrong )
      wire#w1
      { S7_GenerateENO := "TRUE" } Move(in := 3, out1 => #State)
   END_RUNG
   RUNG wire#w1
      S_Coil( #F_RunWrong )
   END_RUNG
   // the same network as SCL:
   IF #RunWrong THEN
       #State := 3;
       #F_RunWrong := TRUE;
   END_IF;
END_REGION

REGION Network 45: E1 / E3 — heat request while STARTING or RUNNING
   RUNG wire#powerrail
      { S7_Templates := "SrcType := Int" } EQ_Contact(in1 := #State, in2 := 1)
      wire#w1
      Coil( #Active )
   END_RUNG
   RUNG wire#powerrail
      { S7_Templates := "SrcType := Int" } EQ_Contact(in1 := #State, in2 := 2)
   END_RUNG wire#w1
   RUNG wire#w1
      Coil( #HeatReq )
   END_RUNG
   // the same network as SCL:
   #Active := (#State = 1) OR (#State = 2);
   #HeatReq := #Active;
END_REGION

REGION Network 46: C0xc — 2nd stage on: RUNNING and T < SP - STG
   RUNG wire#powerrail
      { S7_Templates := "SrcType := Int" } EQ_Contact(in1 := #State, in2 := 2)
      { S7_Templates := "SrcType := Int" } LT_Contact(in1 := #Tmax, in2 := #TStg)
      S_Coil( #Stage2 )
   END_RUNG
   // the same network as SCL:
   IF (#State = 2) AND (#Tmax < #TStg) THEN #Stage2 := TRUE; END_IF;
END_REGION

REGION Network 47: C0xc / F41 — 2nd stage off at SP - STG + 2 degC, or when not RUNNING
   RUNG wire#powerrail
      { S7_Templates := "SrcType := Int" } GE_Contact(in1 := #Tmax, in2 := #TStgOff)
      wire#w1
      R_Coil( #Stage2 )
   END_RUNG
   RUNG wire#powerrail
      { S7_Templates := "SrcType := Int" } NE_Contact(in1 := #State, in2 := 2)
   END_RUNG wire#w1
   // the same network as SCL:
   IF (#Tmax >= #TStgOff) OR (#State <> 2) THEN #Stage2 := FALSE; END_IF;
END_REGION
END_FUNCTION_BLOCK

FUNCTION "Outputs" : Void   // FC2, LAD
TITLE = Outputs
{ S7_Optimized_Access := 'TRUE' }
VERSION : 0.1
// The only block that writes %Q (decisions/0006 rule 3)
// stored: AutoNumber false, IsIECCheckEnabled false, SetENOAutomatically False
BEGIN

REGION Network 1: E1 — BR01 heat request TL (R1, H1)
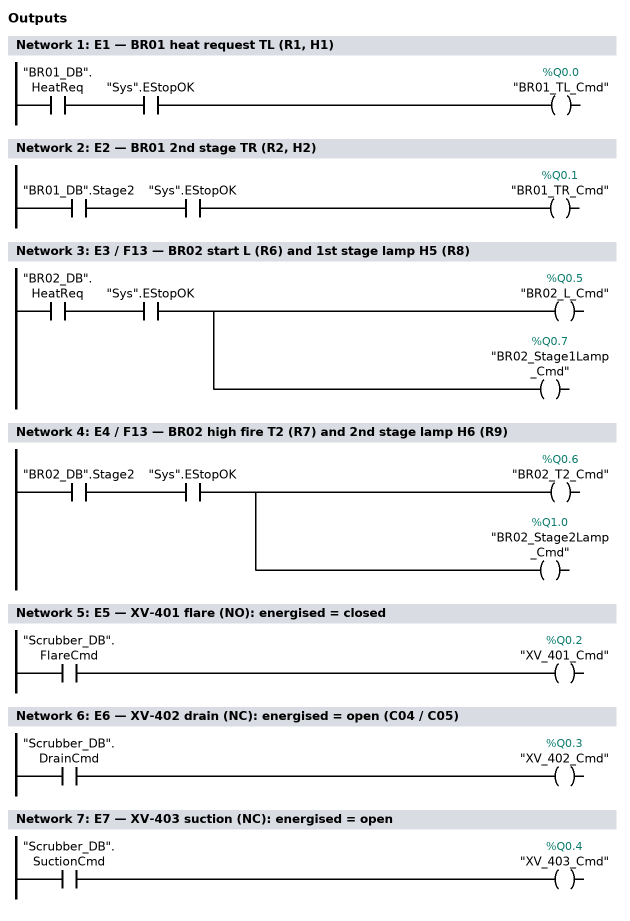
   RUNG wire#powerrail
      Contact( "BR01_DB".HeatReq )
      Contact( "Sys".EStopOK )
      Coil( "BR01_TL_Cmd" )
   END_RUNG
   // the same network as SCL:
   "BR01_TL_Cmd" := "BR01_DB".HeatReq AND "Sys".EStopOK;
END_REGION

REGION Network 2: E2 — BR01 2nd stage TR (R2, H2)
   RUNG wire#powerrail
      Contact( "BR01_DB".Stage2 )
      Contact( "Sys".EStopOK )
      Coil( "BR01_TR_Cmd" )
   END_RUNG
   // the same network as SCL:
   "BR01_TR_Cmd" := "BR01_DB".Stage2 AND "Sys".EStopOK;
END_REGION

REGION Network 3: E3 / F13 — BR02 start L (R6) and 1st stage lamp H5 (R8)
   RUNG wire#powerrail
      Contact( "BR02_DB".HeatReq )
      Contact( "Sys".EStopOK )
      wire#w1
      Coil( "BR02_L_Cmd" )
   END_RUNG
   RUNG wire#w1
      Coil( "BR02_Stage1Lamp_Cmd" )
   END_RUNG
   // the same network as SCL:
   "BR02_L_Cmd" := "BR02_DB".HeatReq AND "Sys".EStopOK;
   "BR02_Stage1Lamp_Cmd" := "BR02_L_Cmd";
END_REGION

REGION Network 4: E4 / F13 — BR02 high fire T2 (R7) and 2nd stage lamp H6 (R9)
   RUNG wire#powerrail
      Contact( "BR02_DB".Stage2 )
      Contact( "Sys".EStopOK )
      wire#w1
      Coil( "BR02_T2_Cmd" )
   END_RUNG
   RUNG wire#w1
      Coil( "BR02_Stage2Lamp_Cmd" )
   END_RUNG
   // the same network as SCL:
   "BR02_T2_Cmd" := "BR02_DB".Stage2 AND "Sys".EStopOK;
   "BR02_Stage2Lamp_Cmd" := "BR02_T2_Cmd";
END_REGION

REGION Network 5: E5 — XV-401 flare (NO): energised = closed
   RUNG wire#powerrail
      Contact( "Scrubber_DB".FlareCmd )
      Coil( "XV_401_Cmd" )
   END_RUNG
   // the same network as SCL:
   "XV_401_Cmd" := "Scrubber_DB".FlareCmd;
END_REGION

REGION Network 6: E6 — XV-402 drain (NC): energised = open (C04 / C05)
   RUNG wire#powerrail
      Contact( "Scrubber_DB".DrainCmd )
      Coil( "XV_402_Cmd" )
   END_RUNG
   // the same network as SCL:
   "XV_402_Cmd" := "Scrubber_DB".DrainCmd;
END_REGION

REGION Network 7: E7 — XV-403 suction (NC): energised = open
   RUNG wire#powerrail
      Contact( "Scrubber_DB".SuctionCmd )
      Coil( "XV_403_Cmd" )
   END_RUNG
   // the same network as SCL:
   "XV_403_Cmd" := "Scrubber_DB".SuctionCmd;
END_REGION
END_FUNCTION

FUNCTION "HmiMap" : Void   // FC3, LAD
TITLE = HmiMap
{ S7_Optimized_Access := 'TRUE' }
VERSION : 0.1
// 0007 / H-05: alarm display map only; writes HmiAlm only, no Ack
// stored: AutoNumber false, IsIECCheckEnabled false, SetENOAutomatically False
BEGIN

REGION Network 1: C01 / 0007 H-05 — Common.x0: E-STOP active or not reset; clears: Release E-STOP and RESET
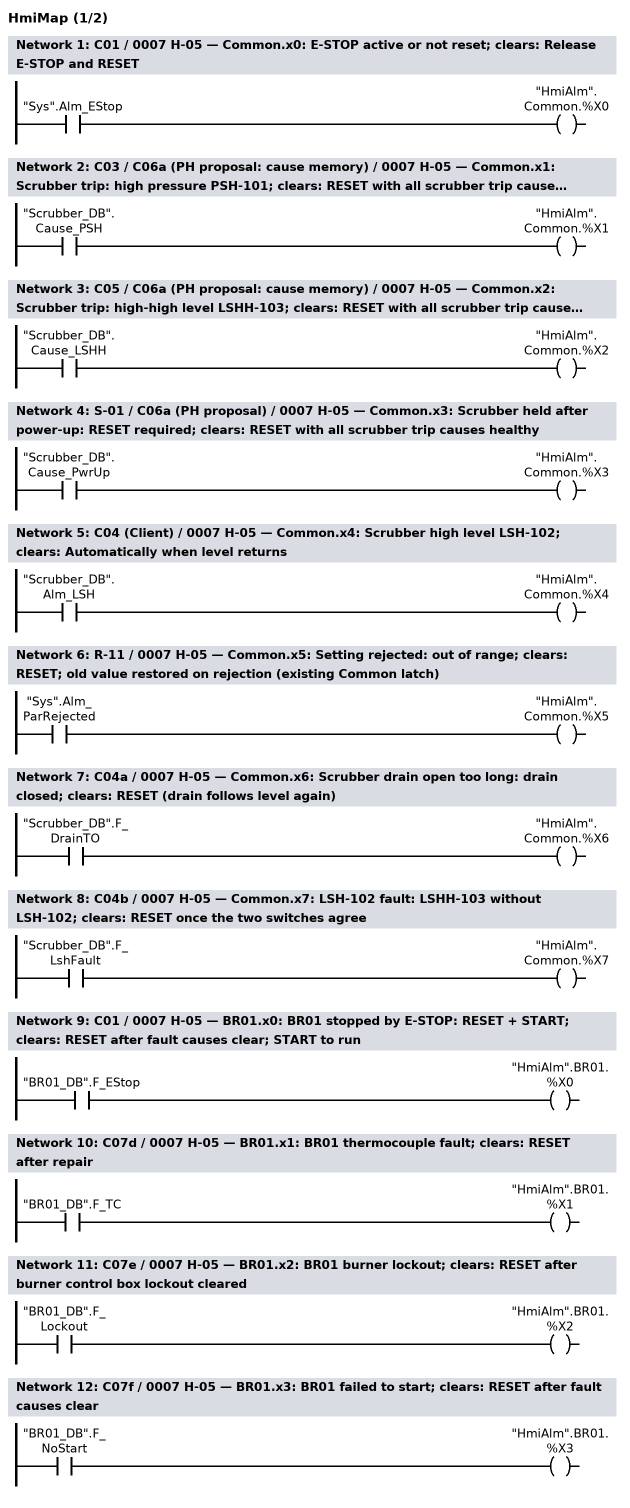
   RUNG wire#powerrail
      Contact( "Sys".Alm_EStop )
      Coil( "HmiAlm".Common.%X0 )
   END_RUNG
   // the same network as SCL:
   "HmiAlm".Common.%X0 := "Sys".Alm_EStop;
END_REGION

REGION Network 2: C03 / C06a (PH proposal: cause memory) / 0007 H-05 — Common.x1: Scrubber trip: high pressure PSH-101; clears: RESET with all scrubber trip causes healthy
   RUNG wire#powerrail
      Contact( "Scrubber_DB".Cause_PSH )
      Coil( "HmiAlm".Common.%X1 )
   END_RUNG
   // the same network as SCL:
   "HmiAlm".Common.%X1 := "Scrubber_DB".Cause_PSH;
END_REGION

REGION Network 3: C05 / C06a (PH proposal: cause memory) / 0007 H-05 — Common.x2: Scrubber trip: high-high level LSHH-103; clears: RESET with all scrubber trip causes healthy
   RUNG wire#powerrail
      Contact( "Scrubber_DB".Cause_LSHH )
      Coil( "HmiAlm".Common.%X2 )
   END_RUNG
   // the same network as SCL:
   "HmiAlm".Common.%X2 := "Scrubber_DB".Cause_LSHH;
END_REGION

REGION Network 4: S-01 / C06a (PH proposal) / 0007 H-05 — Common.x3: Scrubber held after power-up: RESET required; clears: RESET with all scrubber trip causes healthy
   RUNG wire#powerrail
      Contact( "Scrubber_DB".Cause_PwrUp )
      Coil( "HmiAlm".Common.%X3 )
   END_RUNG
   // the same network as SCL:
   "HmiAlm".Common.%X3 := "Scrubber_DB".Cause_PwrUp;
END_REGION

REGION Network 5: C04 (Client) / 0007 H-05 — Common.x4: Scrubber high level LSH-102; clears: Automatically when level returns
   RUNG wire#powerrail
      Contact( "Scrubber_DB".Alm_LSH )
      Coil( "HmiAlm".Common.%X4 )
   END_RUNG
   // the same network as SCL:
   "HmiAlm".Common.%X4 := "Scrubber_DB".Alm_LSH;
END_REGION

REGION Network 6: R-11 / 0007 H-05 — Common.x5: Setting rejected: out of range; clears: RESET; old value restored on rejection (existing Common latch)
   RUNG wire#powerrail
      Contact( "Sys".Alm_ParRejected )
      Coil( "HmiAlm".Common.%X5 )
   END_RUNG
   // the same network as SCL:
   "HmiAlm".Common.%X5 := "Sys".Alm_ParRejected;
END_REGION

REGION Network 7: C04a / 0007 H-05 — Common.x6: Scrubber drain open too long: drain closed; clears: RESET (drain follows level again)
   RUNG wire#powerrail
      Contact( "Scrubber_DB".F_DrainTO )
      Coil( "HmiAlm".Common.%X6 )
   END_RUNG
   // the same network as SCL:
   "HmiAlm".Common.%X6 := "Scrubber_DB".F_DrainTO;
END_REGION

REGION Network 8: C04b / 0007 H-05 — Common.x7: LSH-102 fault: LSHH-103 without LSH-102; clears: RESET once the two switches agree
   RUNG wire#powerrail
      Contact( "Scrubber_DB".F_LshFault )
      Coil( "HmiAlm".Common.%X7 )
   END_RUNG
   // the same network as SCL:
   "HmiAlm".Common.%X7 := "Scrubber_DB".F_LshFault;
END_REGION

REGION Network 9: C01 / 0007 H-05 — BR01.x0: BR01 stopped by E-STOP: RESET + START; clears: RESET after fault causes clear; START to run
   RUNG wire#powerrail
      Contact( "BR01_DB".F_EStop )
      Coil( "HmiAlm".BR01.%X0 )
   END_RUNG
   // the same network as SCL:
   "HmiAlm".BR01.%X0 := "BR01_DB".F_EStop;
END_REGION

REGION Network 10: C07d / 0007 H-05 — BR01.x1: BR01 thermocouple fault; clears: RESET after repair
   RUNG wire#powerrail
      Contact( "BR01_DB".F_TC )
      Coil( "HmiAlm".BR01.%X1 )
   END_RUNG
   // the same network as SCL:
   "HmiAlm".BR01.%X1 := "BR01_DB".F_TC;
END_REGION

REGION Network 11: C07e / 0007 H-05 — BR01.x2: BR01 burner lockout; clears: RESET after burner control box lockout cleared
   RUNG wire#powerrail
      Contact( "BR01_DB".F_Lockout )
      Coil( "HmiAlm".BR01.%X2 )
   END_RUNG
   // the same network as SCL:
   "HmiAlm".BR01.%X2 := "BR01_DB".F_Lockout;
END_REGION

REGION Network 12: C07f / 0007 H-05 — BR01.x3: BR01 failed to start; clears: RESET after fault causes clear
   RUNG wire#powerrail
      Contact( "BR01_DB".F_NoStart )
      Coil( "HmiAlm".BR01.%X3 )
   END_RUNG
   // the same network as SCL:
   "HmiAlm".BR01.%X3 := "BR01_DB".F_NoStart;
END_REGION

REGION Network 13: C07g / 0007 H-05 — BR01.x4: BR01 stopped by itself; clears: RESET after fault causes clear
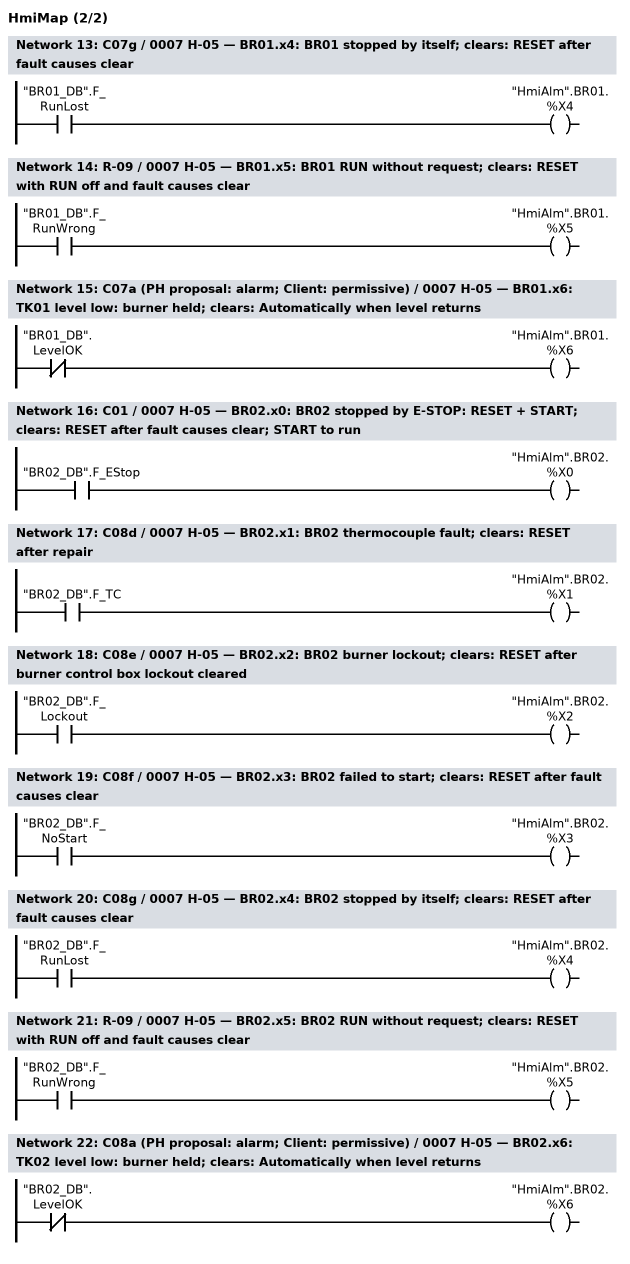
   RUNG wire#powerrail
      Contact( "BR01_DB".F_RunLost )
      Coil( "HmiAlm".BR01.%X4 )
   END_RUNG
   // the same network as SCL:
   "HmiAlm".BR01.%X4 := "BR01_DB".F_RunLost;
END_REGION

REGION Network 14: R-09 / 0007 H-05 — BR01.x5: BR01 RUN without request; clears: RESET with RUN off and fault causes clear
   RUNG wire#powerrail
      Contact( "BR01_DB".F_RunWrong )
      Coil( "HmiAlm".BR01.%X5 )
   END_RUNG
   // the same network as SCL:
   "HmiAlm".BR01.%X5 := "BR01_DB".F_RunWrong;
END_REGION

REGION Network 15: C07a (PH proposal: alarm; Client: permissive) / 0007 H-05 — BR01.x6: TK01 level low: burner held; clears: Automatically when level returns
   RUNG wire#powerrail
      I_Contact( "BR01_DB".LevelOK )
      Coil( "HmiAlm".BR01.%X6 )
   END_RUNG
   // the same network as SCL:
   "HmiAlm".BR01.%X6 := NOT "BR01_DB".LevelOK;
END_REGION

REGION Network 16: C01 / 0007 H-05 — BR02.x0: BR02 stopped by E-STOP: RESET + START; clears: RESET after fault causes clear; START to run
   RUNG wire#powerrail
      Contact( "BR02_DB".F_EStop )
      Coil( "HmiAlm".BR02.%X0 )
   END_RUNG
   // the same network as SCL:
   "HmiAlm".BR02.%X0 := "BR02_DB".F_EStop;
END_REGION

REGION Network 17: C08d / 0007 H-05 — BR02.x1: BR02 thermocouple fault; clears: RESET after repair
   RUNG wire#powerrail
      Contact( "BR02_DB".F_TC )
      Coil( "HmiAlm".BR02.%X1 )
   END_RUNG
   // the same network as SCL:
   "HmiAlm".BR02.%X1 := "BR02_DB".F_TC;
END_REGION

REGION Network 18: C08e / 0007 H-05 — BR02.x2: BR02 burner lockout; clears: RESET after burner control box lockout cleared
   RUNG wire#powerrail
      Contact( "BR02_DB".F_Lockout )
      Coil( "HmiAlm".BR02.%X2 )
   END_RUNG
   // the same network as SCL:
   "HmiAlm".BR02.%X2 := "BR02_DB".F_Lockout;
END_REGION

REGION Network 19: C08f / 0007 H-05 — BR02.x3: BR02 failed to start; clears: RESET after fault causes clear
   RUNG wire#powerrail
      Contact( "BR02_DB".F_NoStart )
      Coil( "HmiAlm".BR02.%X3 )
   END_RUNG
   // the same network as SCL:
   "HmiAlm".BR02.%X3 := "BR02_DB".F_NoStart;
END_REGION

REGION Network 20: C08g / 0007 H-05 — BR02.x4: BR02 stopped by itself; clears: RESET after fault causes clear
   RUNG wire#powerrail
      Contact( "BR02_DB".F_RunLost )
      Coil( "HmiAlm".BR02.%X4 )
   END_RUNG
   // the same network as SCL:
   "HmiAlm".BR02.%X4 := "BR02_DB".F_RunLost;
END_REGION

REGION Network 21: R-09 / 0007 H-05 — BR02.x5: BR02 RUN without request; clears: RESET with RUN off and fault causes clear
   RUNG wire#powerrail
      Contact( "BR02_DB".F_RunWrong )
      Coil( "HmiAlm".BR02.%X5 )
   END_RUNG
   // the same network as SCL:
   "HmiAlm".BR02.%X5 := "BR02_DB".F_RunWrong;
END_REGION

REGION Network 22: C08a (PH proposal: alarm; Client: permissive) / 0007 H-05 — BR02.x6: TK02 level low: burner held; clears: Automatically when level returns
   RUNG wire#powerrail
      I_Contact( "BR02_DB".LevelOK )
      Coil( "HmiAlm".BR02.%X6 )
   END_RUNG
   // the same network as SCL:
   "HmiAlm".BR02.%X6 := NOT "BR02_DB".LevelOK;
END_REGION
END_FUNCTION

ORGANIZATION_BLOCK "Startup"   // OB100, LAD, Startup
TITLE = Startup
{ S7_Optimized_Access := 'TRUE' }
VERSION : 0.1
// Startup OB (decisions/0006)
// stored: AutoNumber false, IsIECCheckEnabled false, SetENOAutomatically False
   VAR_INPUT
      LostRetentive : Bool;
      LostRTC : Bool;
   END_VAR
BEGIN

REGION Network 1: C02 — power-up: first-scan flag (scrubber trips, burners need START)
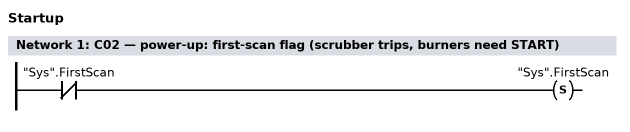
   RUNG wire#powerrail
      I_Contact( "Sys".FirstScan )
      S_Coil( "Sys".FirstScan )
   END_RUNG
   // the same network as SCL:
   IF NOT "Sys".FirstScan THEN "Sys".FirstScan := TRUE; END_IF;
END_REGION
END_ORGANIZATION_BLOCK

DATA_BLOCK "BR01_DB"   // DB3
{ S7_Optimized_Access := 'TRUE' }
VERSION : 0.1
// stored: AutoNumber false, InstanceOfName Burner, InstanceOfType FB
"Burner"
BEGIN
END_DATA_BLOCK

DATA_BLOCK "BR02_DB"   // DB4
{ S7_Optimized_Access := 'TRUE' }
VERSION : 0.1
// stored: AutoNumber false, InstanceOfName Burner, InstanceOfType FB
"Burner"
BEGIN
END_DATA_BLOCK

DATA_BLOCK "Scrubber_DB"   // DB5
{ S7_Optimized_Access := 'TRUE' }
VERSION : 0.1
// stored: AutoNumber false, InstanceOfName Scrubber, InstanceOfType FB
"Scrubber"
BEGIN
END_DATA_BLOCK
